// TIA Portal project "btl" (V17)

(* hardware
DEVICE "S7-1200 station_1"  S7-1200 Station
   slot 0: "Rack_0"  S7-1200 Rack  Rack  V1.0
   slot 1: "PLC_1"  CPU 1215C DC/DC/DC  6ES7 215-1AG40-0XB0  V4.5
   slot 2: "DI 16/DQ 16x24VDC SINK_1"  SM 1223 DI16/DQ16 x 24VDC SINK  6ES7 223-1BL32-1XB0  V2.0
   slot 3: "AI 8x13BIT_1"  6ES7 231-4HF32-0XB0  V2.1
   slot 4: "DI 8x24VDC_1"  SM 1221 DI8 x 24VDC  6ES7 221-1BF30-0XB0  V1.0
DEVICE "PC-System_1"  SIMATIC PC station
   slot 0: "SIMATIC PC station"  Rail  SIMATIC PC-Station  V1.0
      slot 125: "Stationmanager"  Station_Manager  V6.0.4
   slot 1: "HMI_RT_1"  WinCC RT Advanced  6AV2 104-0xxxx-xxxx  17.0.0.0
      slot 33792: "Computer interface"  Host interface
   slot 2: "IE general_1"  IE General  IE_CP  V8.2.0
      slot 1: "PROFINET interface"  IEGeneral.Interface.8.2.0
*)

// ===== PLC "PLC_1"  CPU 1215C DC/DC/DC =====

VAR_GLOBAL   // PLC tag table "Default tag table"
   "System_Byte" AT %MB1 : Byte;
   "FirstScan" AT %M1.0 : Bool;
   "DiagStatusUpdate" AT %M1.1 : Bool;
   "AlwaysTRUE" AT %M1.2 : Bool;
   "AlwaysFALSE" AT %M1.3 : Bool;
   "Clock_Byte" AT %MB0 : Byte;
   "Clock_10Hz" AT %M0.0 : Bool;
   "Clock_5Hz" AT %M0.1 : Bool;
   "Clock_2.5Hz" AT %M0.2 : Bool;
   "Clock_2Hz" AT %M0.3 : Bool;
   "Clock_1.25Hz" AT %M0.4 : Bool;
   "Clock_1Hz" AT %M0.5 : Bool;
   "Clock_0.625Hz" AT %M0.6 : Bool;
   "Clock_0.5Hz" AT %M0.7 : Bool;
END_VAR

VAR_GLOBAL   // PLC tag table "CB_analog"
   "I_Can_huong" AT %IW64 : Int;
   "I_can_mau" AT %IW66 : Int;
   "I_can_Duong" AT %IW68 : Int;
   "I_can_nuoc_TRON" AT %IW70 : Int;
   "I_Can_nuoc_xuc_khi" AT %IW72 : Int;
   "I_Can_PG" AT %IW74 : Int;
   "I_Can_CO2" AT %IW76 : Int;
   "I_bon_1" AT %IW82 : Int;
   "I_bon_2" AT %IW84 : Int;
   "I_bon_3" AT %IW86 : Int;
END_VAR

VAR_GLOBAL   // PLC tag table "INPUT_I"
   "I_mode" AT %I0.0 : Bool;
   "I_start" AT %I0.1 : Bool;
   "I_Stop" AT %I0.2 : Bool;
   "I_SW_V1_Huong" AT %I0.3 : Bool;
   "I_SW_V2_Huong" AT %I0.4 : Bool;
   "I_SW_V1_mau" AT %I0.5 : Bool;
   "I_SW_V2_mau" AT %I0.6 : Bool;
   "I_SW_V1_PG" AT %I0.7 : Bool;
   "I_SW_V2_PG" AT %I1.0 : Bool;
   "I_SW_V1_Duong" AT %I1.1 : Bool;
   "I_SW_V2_Duong" AT %I1.2 : Bool;
   "I_SW_V1_Nuoc_Tron" AT %I1.3 : Bool;
   "I_SW_V2_Nuoc_Tron" AT %I1.4 : Bool;
   "I_SW_V1_Nuoc_Xuc_Khi" AT %I1.5 : Bool;
   "I_SW_V2_Nuoc_Xuc_Khi" AT %I1.6 : Bool;
   "I_SW_V1_CO2" AT %I1.7 : Bool;
   "I_SW_V2_CO2" AT %I2.0 : Bool;
   "I_SW_BOM_TRON" AT %I2.1 : Bool;
   "I_SW_LAM_LANH" AT %I2.2 : Bool;
   "I_SW_BOM_1" AT %I2.3 : Bool;
   "I_SW_BOM_2" AT %I2.4 : Bool;
   "I_SW_LO_DOT" AT %I2.5 : Bool;
   "I_SW_VAN_XA" AT %I2.6 : Bool;
   "I_SW_BANG_TAI" AT %I2.7 : Bool;
   "I_CB_LOW_HUONG" AT %I3.0 : Bool;
   "I_CB_LOW_MAU" AT %I3.1 : Bool;
   "I_CB_LOW_PG" AT %I3.2 : Bool;
   "I_CB_LOW_DUONG" AT %I3.3 : Bool;
   "I_CB_LOW_NUOC" AT %I3.4 : Bool;
   "I_CB_LOW_CO2" AT %I3.5 : Bool;
   "I_CB_CHAI" AT %I3.6 : Bool;
END_VAR

VAR_GLOBAL   // PLC tag table "INPUT_M"
   "M_mode" AT %M10.0 : Bool;
   "M_start" AT %M10.1 : Bool;
   "M_Stop" AT %M10.2 : Bool;
   "M_SW_V1_Huong" AT %M10.3 : Bool;
   "M_SW_V2_Huong" AT %M10.4 : Bool;
   "M_SW_V1_mau" AT %M10.5 : Bool;
   "M_SW_V2_mau" AT %M10.6 : Bool;
   "M_SW_V1_PG" AT %M10.7 : Bool;
   "M_SW_V2_PG" AT %M11.0 : Bool;
   "M_SW_V1_Duong" AT %M11.1 : Bool;
   "M_SW_V2_Duong" AT %M11.2 : Bool;
   "M_SW_V1_Nuoc_Tron" AT %M11.3 : Bool;
   "M_SW_V2_Nuoc_Tron" AT %M11.4 : Bool;
   "M_SW_V1_Nuoc_Xuc_Khi" AT %M11.5 : Bool;
   "M_SW_V2_Nuoc_Xuc_Khi" AT %M11.6 : Bool;
   "M_SW_V1_CO2" AT %M11.7 : Bool;
   "M_SW_V2_CO2" AT %M12.0 : Bool;
   "M_SW_BOM_TRON" AT %M12.1 : Bool;
   "M_SW_LAM_LANH" AT %M12.2 : Bool;
   "M_SW_BOM_1" AT %M12.3 : Bool;
   "M_SW_BOM_2" AT %M12.4 : Bool;
   "M_SW_LO_DOT" AT %M12.5 : Bool;
   "M_SW_VAN_XA" AT %M12.6 : Bool;
   "M_SW_BANG_TAI" AT %M12.7 : Bool;
   "M_CB_LOW_HUONG" AT %M13.0 : Bool;
   "M_CB_LOW_MAU" AT %M13.1 : Bool;
   "M_CB_LOW_PG" AT %M13.2 : Bool;
   "M_CB_LOW_DUONG" AT %M13.3 : Bool;
   "M_CB_LOW_NUOC" AT %M13.4 : Bool;
   "M_CB_LOW_CO2" AT %MD500 : Real;
   "M_CB_LOW_BON_2" AT %MD504 : Real;
   "M_CB_CHAI" AT %M13.7 : Bool;
END_VAR

VAR_GLOBAL   // PLC tag table "OUTPUT"
   "Q_den_Auto" AT %Q0.0 : Bool;
   "Q_Den_Manual" AT %Q0.1 : Bool;
   "Q_Den_loi" AT %Q0.2 : Bool;
   "Q_V1_Huong" AT %Q0.3 : Bool;
   "Q_V2_Huong" AT %Q0.4 : Bool;
   "Q_V1_Mau" AT %Q0.5 : Bool;
   "Q_V2_Mau" AT %Q0.6 : Bool;
   "Q_V1_PG" AT %Q0.7 : Bool;
   "Q_V2_PG" AT %Q1.0 : Bool;
   "Q_V1_Nuoc_Tron" AT %Q1.1 : Bool;
   "Q_V2_Nuoc_tron" AT %Q1.2 : Bool;
   "Q_V1_Duong" AT %Q1.3 : Bool;
   "Q_V2_Duong" AT %Q1.4 : Bool;
   "Q_V1_Nuoc_Khi" AT %Q1.5 : Bool;
   "Q_V2_Xuc_Khi" AT %Q1.6 : Bool;
   "Q_V1_CO2" AT %Q1.7 : Bool;
   "Q_V2_CO2" AT %Q2.0 : Bool;
   "Q_BOM_TRON" AT %Q2.1 : Bool;
   "Q_LAM_LANH" AT %Q2.2 : Bool;
   "Q_BOM_1" AT %Q2.3 : Bool;
   "Q_BOM_2" AT %Q2.4 : Bool;
   "Q_VAN_XA" AT %Q2.5 : Bool;
   "Q_LO_DOT" AT %Q2.6 : Bool;
   "Q_BT" AT %Q2.7 : Bool;
END_VAR

VAR_GLOBAL   // PLC tag table "OUTPUT_AUTO"
   "Q_AUTO_den_Auto" AT %M20.0 : Bool;
   "Q_AUTO_Den_Manual" AT %M20.1 : Bool;
   "Q_AUTO_Den_loi" AT %M20.2 : Bool;
   "Q_AUTO_V1_Huong" AT %M20.3 : Bool;
   "Q_AUTO_V2_Huong" AT %M20.4 : Bool;
   "Q_AUTO_V1_Mau" AT %M20.5 : Bool;
   "Q_AUTO_V2_Mau" AT %M20.6 : Bool;
   "Q_AUTO_V1_PG" AT %M20.7 : Bool;
   "Q_AUTO_V2_PG" AT %M21.0 : Bool;
   "Q_AUTO_V1_Nuoc_Tron" AT %M21.1 : Bool;
   "Q_AUTO_V2_Nuoc_tron" AT %M21.2 : Bool;
   "Q_AUTO_V1_Duong" AT %M21.3 : Bool;
   "Q_AUTO_V2_Duong" AT %M21.4 : Bool;
   "Q_AUTO_V1_Nuoc_Khi" AT %M21.5 : Bool;
   "Q_AUTO_V2_Xuc_Khi" AT %M21.6 : Bool;
   "Q_AUTO_V1_CO2" AT %M21.7 : Bool;
   "Q_AUTO_V2_CO2" AT %M22.0 : Bool;
   "Q_AUTO_BOM_TRON" AT %M22.1 : Bool;
   "Q_AUTO_LAM_LANH" AT %M22.2 : Bool;
   "Q_AUTO_BOM_1" AT %M22.3 : Bool;
   "Q_AUTO_BOM_2" AT %M22.4 : Bool;
   "Q_AUTO_VAN_XA" AT %M22.5 : Bool;
   "Q_AUTO_LO_DOT" AT %M22.6 : Bool;
   "Q_AUTO_BT" AT %M22.7 : Bool;
END_VAR

VAR_GLOBAL   // PLC tag table "OUTPUT_MANUAL"
   "Q_MAN_den_Auto" AT %M30.0 : Bool;
   "Q_MAN_Den_Manual" AT %M30.1 : Bool;
   "Q_MAN_Den_loi" AT %M30.2 : Bool;
   "Q_MAN_V1_Huong" AT %M30.3 : Bool;
   "Q_MAN_V2_Huong" AT %M30.4 : Bool;
   "Q_MAN_V1_Mau" AT %M30.5 : Bool;
   "Q_MAN_V2_Mau" AT %M30.6 : Bool;
   "Q_MAN_V1_PG" AT %M30.7 : Bool;
   "Q_MAN_V2_PG" AT %M31.0 : Bool;
   "Q_MAN_V1_Nuoc_Tron" AT %M31.1 : Bool;
   "Q_MAN_V2_Nuoc_tron" AT %M31.2 : Bool;
   "Q_MAN_V1_Duong" AT %M31.3 : Bool;
   "Q_MAN_V2_Duong" AT %M31.4 : Bool;
   "Q_MAN_V1_Nuoc_Khi" AT %M31.5 : Bool;
   "Q_MAN_V2_Xuc_Khi" AT %M31.6 : Bool;
   "Q_MAN_V1_CO2" AT %M31.7 : Bool;
   "Q_MAN_V2_CO2" AT %M32.0 : Bool;
   "Q_MAN_BOM_TRON" AT %M32.1 : Bool;
   "Q_MAN_LAM_LANH" AT %M32.2 : Bool;
   "Q_MAN_BOM_1" AT %M32.3 : Bool;
   "Q_MAN_BOM_2" AT %M32.4 : Bool;
   "Q_MAN_VAN_XA" AT %M32.5 : Bool;
   "Q_MAN_LO_DOT" AT %M32.6 : Bool;
   "Q_MAN_BT" AT %M32.7 : Bool;
END_VAR

VAR_GLOBAL   // PLC tag table "GT_Thuc_TE"
   "Act_time_Khuay" AT %MW400 : Int;
   "Act_nhiet_do" AT %MD402 : Real;
   "Act_me" AT %MW406 : Int;
   "Act_can_huong" AT %MD408 : Real;
   "Act_can_mau" AT %MD412 : Real;
   "Act_can_duong" AT %MD416 : Real;
   "Act_can_PG" AT %MD420 : Real;
   "Act_can_nuoc_tron" AT %MD424 : Real;
   "Act_can_nuoc_xuc_khi" AT %MD428 : Real;
   "Act_Can_CO2" AT %MD432 : Real;
   "Act_So_chai" AT %MW436 : Int;
   "Act_bon_1" AT %MD440 : Real;
   "Act_bon_2" AT %MD444 : Real;
   "Act_bon_3" AT %MD448 : Real;
END_VAR

VAR_GLOBAL   // PLC tag table "Trung_gian"
   "TG_Button_Simulation" AT %M40.0 : Bool;
   "TG_Step_1" AT %M40.1 : Bool;
   "TG_Step_2" AT %M40.2 : Bool;
   "TG_Step_3" AT %M40.3 : Bool;
   "TG_Step_4" AT %M40.4 : Bool;
   "TG_Step_5" AT %M40.5 : Bool;
   "TG_Step_6" AT %M40.6 : Bool;
   "TG_Step_7" AT %M40.7 : Bool;
   "TG_DK_RUN" AT %M41.0 : Bool;
   "TG_Lap_lai" AT %M41.1 : Bool;
   "TG_Can_Xong_huong" AT %M41.2 : Bool;
   "TG_Xung_100ms" AT %M41.3 : Bool;
   "TG_Can_Xong_mau" AT %M41.4 : Bool;
   "TG_Can_Xong_PG" AT %M41.5 : Bool;
   "TG_can_Xong_Nuoc_Khi" AT %M41.6 : Bool;
   "TG_Can_Xong_CO2" AT %M41.7 : Bool;
   "TG_xong_nuoc_tron" AT %M42.0 : Bool;
   "TG_Xong_Nuoc_khi" AT %M42.1 : Bool;
   "TG_xong_huong" AT %M42.2 : Bool;
   "TG_Xong_mau" AT %M42.3 : Bool;
   "TG_Xong_PG" AT %M42.4 : Bool;
   "TG_Xong_duong" AT %M42.5 : Bool;
   "TG_Xong_CO2" AT %M42.6 : Bool;
   "TG_Xong_Khuay" AT %M42.7 : Bool;
   "TG_Xong_Dot" AT %M43.0 : Bool;
   "TG_Thoi_Gian_Dong_SP" AT %M43.1 : Bool;
   "TG_XONG_BANG_TAI" AT %M43.2 : Bool;
   "TG_DONE_CHU_TRINH" AT %M43.3 : Bool;
   "TG_VT_SP" AT %MD508 : DInt;
   "TG_TG_SP" AT %MD512 : DInt;
   "TG_Can_huong" AT %MD516 : Real;
   "TG_Can_mau" AT %MD520 : Real;
   "TG_Can_PG" AT %MD524 : Real;
   "TG_CAn_Duong" AT %MD528 : Real;
   "TG_Can_nuoc_tron" AT %MD532 : Real;
   "TG_Can_nuoc_khi" AT %MD536 : Real;
   "TG_Can_CO2" AT %MD540 : Real;
   "TG_BON1" AT %M43.4 : Bool;
   "TG_BON2" AT %M43.5 : Bool;
   "TG_BON3" AT %M43.6 : Bool;
   "TG_V_BON1" AT %MD544 : Real;
   "TG_V_BON2" AT %MD548 : Real;
   "TG_V_BON3" AT %MD552 : Real;
   "TG_LO_DOT" AT %M43.7 : Bool;
END_VAR

VAR_GLOBAL   // PLC tag table "Trung_giang_Xung"
   "P1" AT %M50.0 : Bool;
   "P2" AT %M50.1 : Bool;
   "P3" AT %M50.2 : Bool;
   "P4" AT %M50.3 : Bool;
   "P5" AT %M50.4 : Bool;
   "P6" AT %M50.5 : Bool;
   "P7" AT %M50.6 : Bool;
   "P8" AT %M50.7 : Bool;
   "P9" AT %M51.0 : Bool;
   "P10" AT %M51.1 : Bool;
   "P11" AT %M51.2 : Bool;
   "P12" AT %M51.3 : Bool;
   "P13" AT %M51.4 : Bool;
   "P14" AT %M51.5 : Bool;
   "P15" AT %M51.6 : Bool;
   "P16" AT %M51.7 : Bool;
   "P17" AT %M52.0 : Bool;
   "P18" AT %M52.1 : Bool;
   "P19" AT %M52.2 : Bool;
   "P20" AT %M52.3 : Bool;
   "P21" AT %M52.4 : Bool;
   "P22" AT %M52.5 : Bool;
   "P23" AT %M52.6 : Bool;
   "P24" AT %M52.7 : Bool;
   "P25" AT %M53.0 : Bool;
   "P26" AT %M53.1 : Bool;
   "P27" AT %M53.2 : Bool;
   "P28" AT %M53.3 : Bool;
   "P29" AT %M53.4 : Bool;
   "P30" AT %M53.5 : Bool;
   "P31" AT %M53.6 : Bool;
   "P32" AT %M53.7 : Bool;
   "P33" AT %M54.0 : Bool;
   "P34" AT %M54.1 : Bool;
   "P35" AT %M54.2 : Bool;
   "P36" AT %M54.3 : Bool;
   "P37" AT %M54.4 : Bool;
   "P38" AT %M54.5 : Bool;
   "P39" AT %M54.6 : Bool;
   "P40" AT %M54.7 : Bool;
   "P41" AT %M55.0 : Bool;
   "P42" AT %M55.1 : Bool;
END_VAR

VAR_GLOBAL   // PLC tag table "Setting"
   "Set_can_huong" AT %MD200 : Real;
   "Set_can_mau" AT %MD204 : Real;
   "Set_can_PG" AT %MD208 : Real;
   "Set_can_Duong" AT %MD212 : Real;
   "Set_Can_nuoc_Tron" AT %MD216 : Real;
   "Set_Can_nuoc_xuc_khi" AT %MD220 : Real;
   "Set_Can_CO2" AT %MD224 : Real;
   "Set_thoi_gian_khuay" AT %MW228 : Int;
   "Set_nhiet_do" AT %MD300 : Real;
   "Set_me_tron" AT %MW304 : Int;
END_VAR

VAR_GLOBAL   // PLC tag table "TRONG LUONG DAT DUOC"
   "TL_Huong" AT %MD600 : Real;
   "TL_mau" AT %MD604 : Real;
   "TL_Duong" AT %MD608 : Real;
   "TL_PG" AT %MD612 : Real;
   "TL_nuoc_tron" AT %MD616 : Real;
   "TL_CO2" AT %MD620 : Real;
   "TL_Nuoc_KHi" AT %MD624 : Real;
   "TL_San_Pham" AT %MD628 : Real;
   "TL_thoiGian_khuay" AT %MD632 : DInt;
   "TL_nhietdo" AT %MD636 : Real;
END_VAR

// folder: System blocks/Program resources

DATA_BLOCK "IEC_Timer_0_DB"   // DB1
{ S7_Optimized_Access := 'TRUE' }
AUTHOR : Simatic
FAMILY : IEC
NAME : IEC_TMR
VERSION : 1.0
// stored: InstanceOfName IEC_TIMER
"IEC_TIMER"
BEGIN
END_DATA_BLOCK

DATA_BLOCK "IEC_Timer_0_DB_1"   // DB2
{ S7_Optimized_Access := 'TRUE' }
AUTHOR : Simatic
FAMILY : IEC
NAME : IEC_TMR
VERSION : 1.0
// stored: InstanceOfName IEC_TIMER
"IEC_TIMER"
BEGIN
END_DATA_BLOCK

DATA_BLOCK "IEC_Timer_0_DB_2"   // DB3
{ S7_Optimized_Access := 'TRUE' }
AUTHOR : Simatic
FAMILY : IEC
NAME : IEC_TMR
VERSION : 1.0
// stored: InstanceOfName IEC_TIMER
"IEC_TIMER"
BEGIN
END_DATA_BLOCK

DATA_BLOCK "IEC_Timer_0_DB_3"   // DB4
{ S7_Optimized_Access := 'TRUE' }
AUTHOR : Simatic
FAMILY : IEC
NAME : IEC_TMR
VERSION : 1.0
// stored: InstanceOfName IEC_TIMER
"IEC_TIMER"
BEGIN
END_DATA_BLOCK

// folder: (top level)

FUNCTION "FC_ANALOG" : Void   // FC1, LAD
{ S7_Optimized_Access := 'TRUE' }
VERSION : 0.1
BEGIN

REGION Network 1: Can Huong
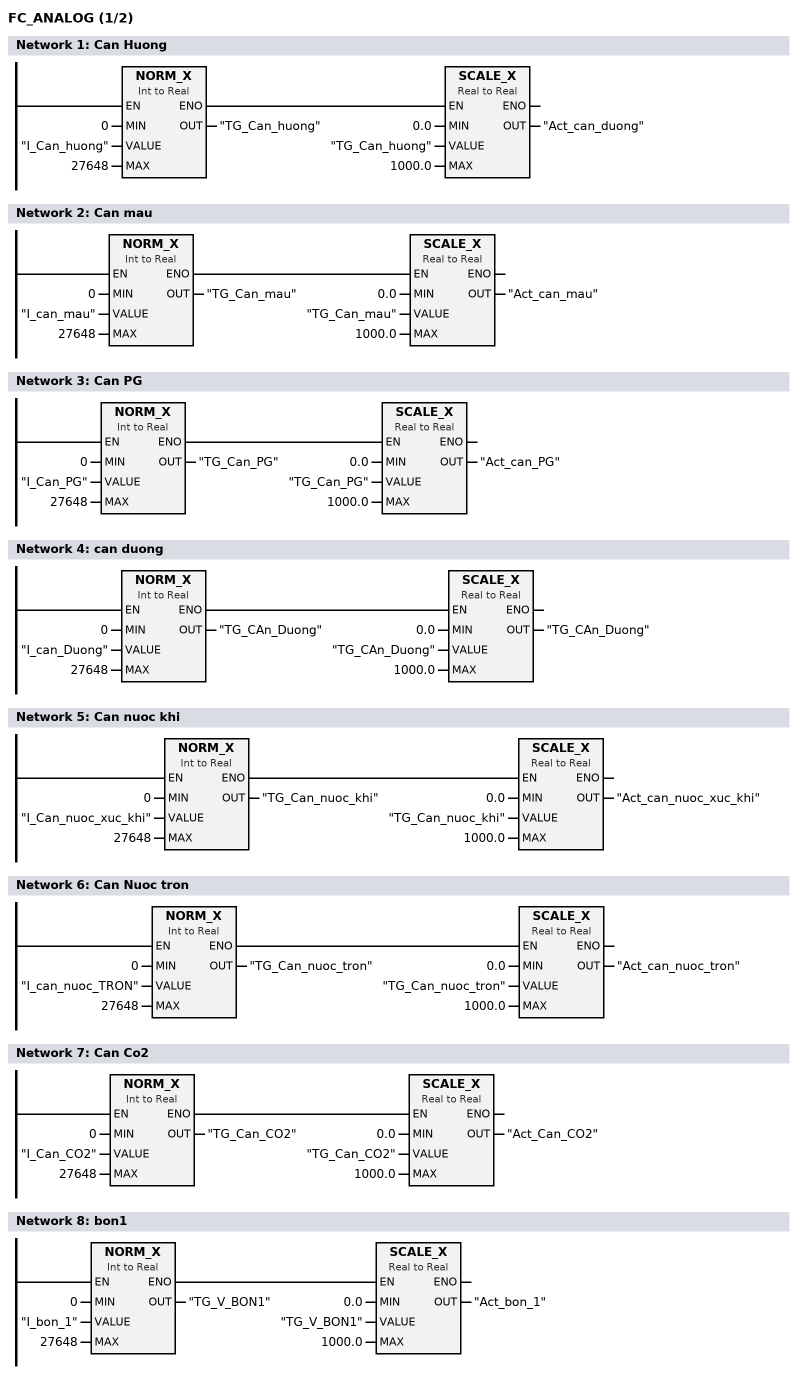
   RUNG wire#powerrail
      { S7_Templates := "[SrcType := Int, DestType := Real]" } Normalize(min := 0, value := "I_Can_huong", max := 27648, out => "TG_Can_huong")
      { S7_Templates := "[SrcType := Real, DestType := Real]" } Scale(min := 0.0, value := "TG_Can_huong", max := 1000.0, out => "Act_can_duong")
   END_RUNG
   // the same network as SCL:
   "TG_Can_huong" := NORM_X(MIN := 0, VALUE := "I_Can_huong", MAX := 27648);
   "Act_can_duong" := SCALE_X(MIN := 0.0, VALUE := "TG_Can_huong", MAX := 1000.0);
END_REGION

REGION Network 2: Can mau
   RUNG wire#powerrail
      { S7_Templates := "[SrcType := Int, DestType := Real]" } Normalize(min := 0, value := "I_can_mau", max := 27648, out => "TG_Can_mau")
      { S7_Templates := "[SrcType := Real, DestType := Real]" } Scale(min := 0.0, value := "TG_Can_mau", max := 1000.0, out => "Act_can_mau")
   END_RUNG
   // the same network as SCL:
   "TG_Can_mau" := NORM_X(MIN := 0, VALUE := "I_can_mau", MAX := 27648);
   "Act_can_mau" := SCALE_X(MIN := 0.0, VALUE := "TG_Can_mau", MAX := 1000.0);
END_REGION

REGION Network 3: Can PG
   RUNG wire#powerrail
      { S7_Templates := "[SrcType := Int, DestType := Real]" } Normalize(min := 0, value := "I_Can_PG", max := 27648, out => "TG_Can_PG")
      { S7_Templates := "[SrcType := Real, DestType := Real]" } Scale(min := 0.0, value := "TG_Can_PG", max := 1000.0, out => "Act_can_PG")
   END_RUNG
   // the same network as SCL:
   "TG_Can_PG" := NORM_X(MIN := 0, VALUE := "I_Can_PG", MAX := 27648);
   "Act_can_PG" := SCALE_X(MIN := 0.0, VALUE := "TG_Can_PG", MAX := 1000.0);
END_REGION

REGION Network 4: can duong
   RUNG wire#powerrail
      { S7_Templates := "[SrcType := Int, DestType := Real]" } Normalize(min := 0, value := "I_can_Duong", max := 27648, out => "TG_CAn_Duong")
      { S7_Templates := "[SrcType := Real, DestType := Real]" } Scale(min := 0.0, value := "TG_CAn_Duong", max := 1000.0, out => "TG_CAn_Duong")
   END_RUNG
   // the same network as SCL:
   "TG_CAn_Duong" := NORM_X(MIN := 0, VALUE := "I_can_Duong", MAX := 27648);
   "TG_CAn_Duong" := SCALE_X(MIN := 0.0, VALUE := "TG_CAn_Duong", MAX := 1000.0);
END_REGION

REGION Network 5: Can nuoc khi
   RUNG wire#powerrail
      { S7_Templates := "[SrcType := Int, DestType := Real]" } Normalize(min := 0, value := "I_Can_nuoc_xuc_khi", max := 27648, out => "TG_Can_nuoc_khi")
      { S7_Templates := "[SrcType := Real, DestType := Real]" } Scale(min := 0.0, value := "TG_Can_nuoc_khi", max := 1000.0, out => "Act_can_nuoc_xuc_khi")
   END_RUNG
   // the same network as SCL:
   "TG_Can_nuoc_khi" := NORM_X(MIN := 0, VALUE := "I_Can_nuoc_xuc_khi", MAX := 27648);
   "Act_can_nuoc_xuc_khi" := SCALE_X(MIN := 0.0, VALUE := "TG_Can_nuoc_khi", MAX := 1000.0);
END_REGION

REGION Network 6: Can Nuoc tron
   RUNG wire#powerrail
      { S7_Templates := "[SrcType := Int, DestType := Real]" } Normalize(min := 0, value := "I_can_nuoc_TRON", max := 27648, out => "TG_Can_nuoc_tron")
      { S7_Templates := "[SrcType := Real, DestType := Real]" } Scale(min := 0.0, value := "TG_Can_nuoc_tron", max := 1000.0, out => "Act_can_nuoc_tron")
   END_RUNG
   // the same network as SCL:
   "TG_Can_nuoc_tron" := NORM_X(MIN := 0, VALUE := "I_can_nuoc_TRON", MAX := 27648);
   "Act_can_nuoc_tron" := SCALE_X(MIN := 0.0, VALUE := "TG_Can_nuoc_tron", MAX := 1000.0);
END_REGION

REGION Network 7: Can Co2
   RUNG wire#powerrail
      { S7_Templates := "[SrcType := Int, DestType := Real]" } Normalize(min := 0, value := "I_Can_CO2", max := 27648, out => "TG_Can_CO2")
      { S7_Templates := "[SrcType := Real, DestType := Real]" } Scale(min := 0.0, value := "TG_Can_CO2", max := 1000.0, out => "Act_Can_CO2")
   END_RUNG
   // the same network as SCL:
   "TG_Can_CO2" := NORM_X(MIN := 0, VALUE := "I_Can_CO2", MAX := 27648);
   "Act_Can_CO2" := SCALE_X(MIN := 0.0, VALUE := "TG_Can_CO2", MAX := 1000.0);
END_REGION

REGION Network 8: bon1
   RUNG wire#powerrail
      { S7_Templates := "[SrcType := Int, DestType := Real]" } Normalize(min := 0, value := "I_bon_1", max := 27648, out => "TG_V_BON1")
      { S7_Templates := "[SrcType := Real, DestType := Real]" } Scale(min := 0.0, value := "TG_V_BON1", max := 1000.0, out => "Act_bon_1")
   END_RUNG
   // the same network as SCL:
   "TG_V_BON1" := NORM_X(MIN := 0, VALUE := "I_bon_1", MAX := 27648);
   "Act_bon_1" := SCALE_X(MIN := 0.0, VALUE := "TG_V_BON1", MAX := 1000.0);
END_REGION

REGION Network 9: bon2
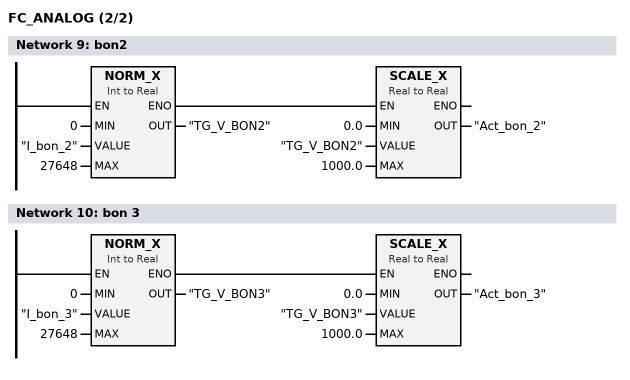
   RUNG wire#powerrail
      { S7_Templates := "[SrcType := Int, DestType := Real]" } Normalize(min := 0, value := "I_bon_2", max := 27648, out => "TG_V_BON2")
      { S7_Templates := "[SrcType := Real, DestType := Real]" } Scale(min := 0.0, value := "TG_V_BON2", max := 1000.0, out => "Act_bon_2")
   END_RUNG
   // the same network as SCL:
   "TG_V_BON2" := NORM_X(MIN := 0, VALUE := "I_bon_2", MAX := 27648);
   "Act_bon_2" := SCALE_X(MIN := 0.0, VALUE := "TG_V_BON2", MAX := 1000.0);
END_REGION

REGION Network 10: bon 3
   RUNG wire#powerrail
      { S7_Templates := "[SrcType := Int, DestType := Real]" } Normalize(min := 0, value := "I_bon_3", max := 27648, out => "TG_V_BON3")
      { S7_Templates := "[SrcType := Real, DestType := Real]" } Scale(min := 0.0, value := "TG_V_BON3", max := 1000.0, out => "Act_bon_3")
   END_RUNG
   // the same network as SCL:
   "TG_V_BON3" := NORM_X(MIN := 0, VALUE := "I_bon_3", MAX := 27648);
   "Act_bon_3" := SCALE_X(MIN := 0.0, VALUE := "TG_V_BON3", MAX := 1000.0);
END_REGION
END_FUNCTION

FUNCTION "FC_AUTO" : Void   // FC2, LAD
{ S7_Optimized_Access := 'TRUE' }
VERSION : 0.1
   VAR_TEMP   // added for the SCL form of the ladder/FBD networks
      _w1 : Bool;
      _w2 : Bool;
      _w3 : Bool;
      _w4 : Bool;
      _w5 : Bool;
      _w6 : Bool;
      _w7 : Bool;
      _w8 : Bool;
      _w9 : Bool;
      _w10 : Bool;
      _w11 : Bool;
      _w12 : Bool;
      _w13 : Bool;
      _w14 : Bool;
      _w15 : Bool;
      _w16 : Bool;
      _w17 : Bool;
      _w18 : Bool;
      _w19 : Bool;
      _w20 : Bool;
      _w21 : Bool;
   END_VAR
BEGIN

REGION Network 1: Điều Kiện Vận Hành
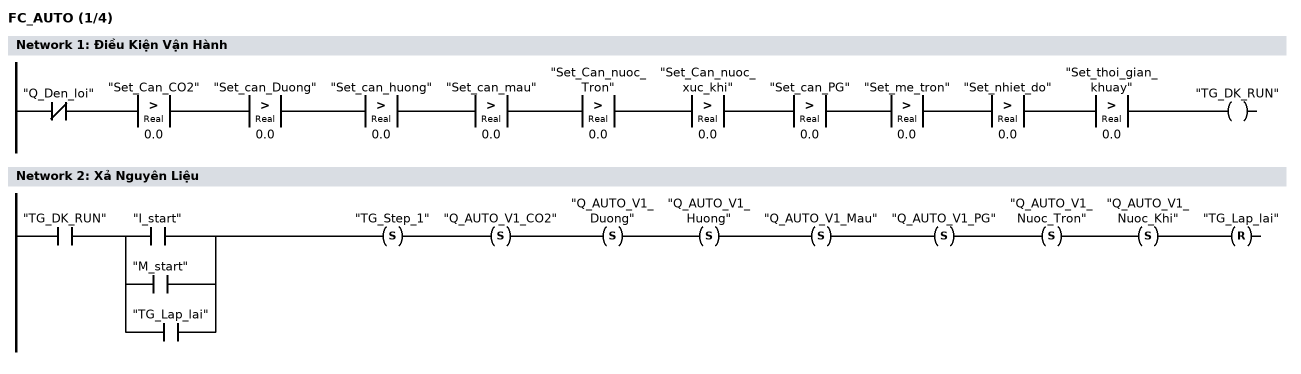
   RUNG wire#powerrail
      I_Contact( "Q_Den_loi" )
      { S7_Templates := "SrcType := Real" } GT_Contact(in1 := "Set_Can_CO2", in2 := 0.0)
      { S7_Templates := "SrcType := Real" } GT_Contact(in1 := "Set_can_Duong", in2 := 0.0)
      { S7_Templates := "SrcType := Real" } GT_Contact(in1 := "Set_can_huong", in2 := 0.0)
      { S7_Templates := "SrcType := Real" } GT_Contact(in1 := "Set_can_mau", in2 := 0.0)
      { S7_Templates := "SrcType := Real" } GT_Contact(in1 := "Set_Can_nuoc_Tron", in2 := 0.0)
      { S7_Templates := "SrcType := Real" } GT_Contact(in1 := "Set_Can_nuoc_xuc_khi", in2 := 0.0)
      { S7_Templates := "SrcType := Real" } GT_Contact(in1 := "Set_can_PG", in2 := 0.0)
      { S7_Templates := "SrcType := Real" } GT_Contact(in1 := "Set_me_tron", in2 := 0.0)
      { S7_Templates := "SrcType := Real" } GT_Contact(in1 := "Set_nhiet_do", in2 := 0.0)
      { S7_Templates := "SrcType := Real" } GT_Contact(in1 := "Set_thoi_gian_khuay", in2 := 0.0)
      Coil( "TG_DK_RUN" )
   END_RUNG
   // the same network as SCL:
   "TG_DK_RUN" := NOT "Q_Den_loi" AND ("Set_Can_CO2" > 0.0) AND ("Set_can_Duong" > 0.0) AND ("Set_can_huong" > 0.0) AND ("Set_can_mau" > 0.0) AND ("Set_Can_nuoc_Tron" > 0.0) AND ("Set_Can_nuoc_xuc_khi" > 0.0) AND ("Set_can_PG" > 0.0) AND ("Set_me_tron" > 0.0) AND ("Set_nhiet_do" > 0.0) AND ("Set_thoi_gian_khuay" > 0.0);
END_REGION

REGION Network 2: Xả Nguyên Liệu
   RUNG wire#powerrail
      Contact( "TG_DK_RUN" )
      wire#w1
      Contact( "I_start" )
      wire#w2
      S_Coil( "TG_Step_1" )
      S_Coil( "Q_AUTO_V1_CO2" )
      S_Coil( "Q_AUTO_V1_Duong" )
      S_Coil( "Q_AUTO_V1_Huong" )
      S_Coil( "Q_AUTO_V1_Mau" )
      S_Coil( "Q_AUTO_V1_PG" )
      S_Coil( "Q_AUTO_V1_Nuoc_Tron" )
      S_Coil( "Q_AUTO_V1_Nuoc_Khi" )
      R_Coil( "TG_Lap_lai" )
   END_RUNG
   RUNG wire#w1
      Contact( "M_start" )
   END_RUNG wire#w2
   RUNG wire#w1
      Contact( "TG_Lap_lai" )
   END_RUNG wire#w2
   // the same network as SCL:
   IF "TG_DK_RUN" AND ("I_start" OR "M_start" OR "TG_Lap_lai") THEN
       "TG_Step_1" := TRUE;
       "Q_AUTO_V1_CO2" := TRUE;
       "Q_AUTO_V1_Duong" := TRUE;
       "Q_AUTO_V1_Huong" := TRUE;
       "Q_AUTO_V1_Mau" := TRUE;
       "Q_AUTO_V1_PG" := TRUE;
       "Q_AUTO_V1_Nuoc_Tron" := TRUE;
       "Q_AUTO_V1_Nuoc_Khi" := TRUE;
       "TG_Lap_lai" := FALSE;
   END_IF;
END_REGION

REGION Network 3: Cân Hương, Đường, Màu , Phụ Gia , Nước , CO2
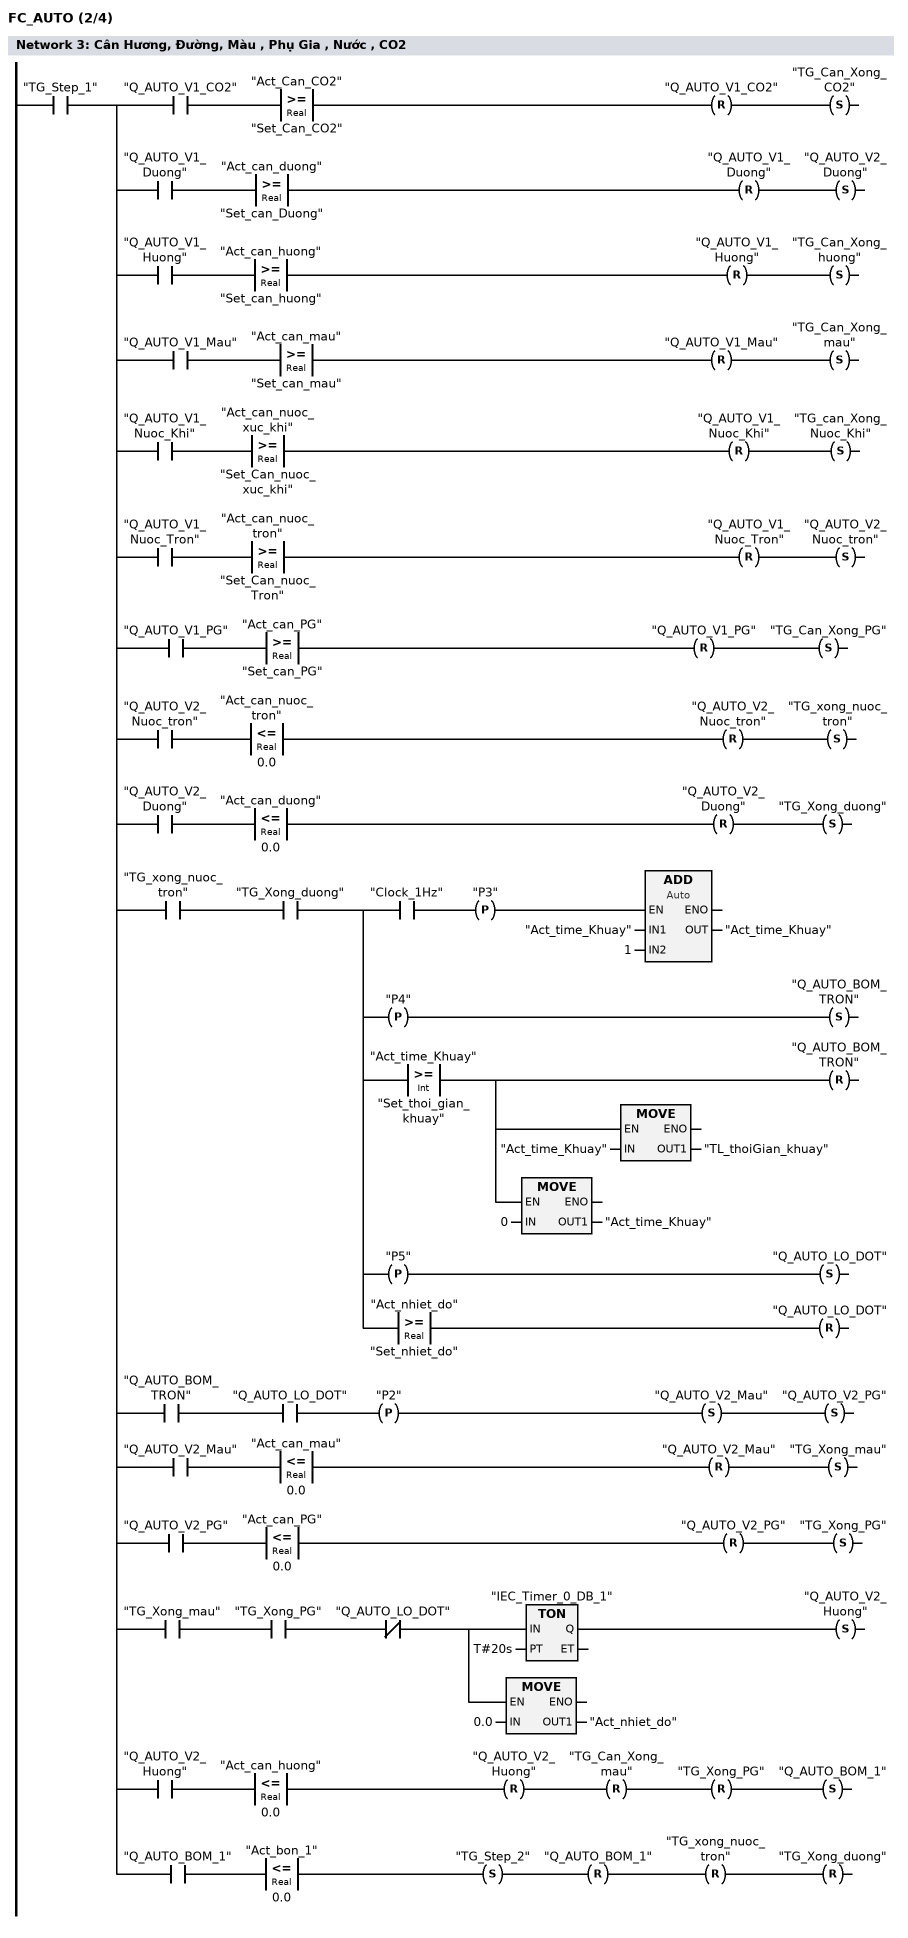
   #_w1 := "TG_Step_1" AND "Q_AUTO_V1_CO2" AND ("Act_Can_CO2" >= "Set_Can_CO2");
   IF #_w1 THEN
       "Q_AUTO_V1_CO2" := FALSE;
       "TG_Can_Xong_CO2" := TRUE;
   END_IF;
   #_w2 := "TG_Step_1" AND "Q_AUTO_V1_Duong" AND ("Act_can_duong" >= "Set_can_Duong");
   IF #_w2 THEN
       "Q_AUTO_V1_Duong" := FALSE;
       "Q_AUTO_V2_Duong" := TRUE;
   END_IF;
   #_w3 := "TG_Step_1" AND "Q_AUTO_V1_Huong" AND ("Act_can_huong" >= "Set_can_huong");
   IF #_w3 THEN
       "Q_AUTO_V1_Huong" := FALSE;
       "TG_Can_Xong_huong" := TRUE;
   END_IF;
   #_w4 := "TG_Step_1" AND "Q_AUTO_V1_Mau" AND ("Act_can_mau" >= "Set_can_mau");
   IF #_w4 THEN
       "Q_AUTO_V1_Mau" := FALSE;
       "TG_Can_Xong_mau" := TRUE;
   END_IF;
   #_w5 := "TG_Step_1" AND "Q_AUTO_V1_Nuoc_Khi" AND ("Act_can_nuoc_xuc_khi" >= "Set_Can_nuoc_xuc_khi");
   IF #_w5 THEN
       "Q_AUTO_V1_Nuoc_Khi" := FALSE;
       "TG_can_Xong_Nuoc_Khi" := TRUE;
   END_IF;
   #_w6 := "TG_Step_1" AND "Q_AUTO_V1_Nuoc_Tron" AND ("Act_can_nuoc_tron" >= "Set_Can_nuoc_Tron");
   IF #_w6 THEN
       "Q_AUTO_V1_Nuoc_Tron" := FALSE;
       "Q_AUTO_V2_Nuoc_tron" := TRUE;
   END_IF;
   #_w7 := "TG_Step_1" AND "Q_AUTO_V1_PG" AND ("Act_can_PG" >= "Set_can_PG");
   IF #_w7 THEN
       "Q_AUTO_V1_PG" := FALSE;
       "TG_Can_Xong_PG" := TRUE;
   END_IF;
   #_w8 := "TG_Step_1" AND "Q_AUTO_V2_Nuoc_tron" AND ("Act_can_nuoc_tron" <= 0.0);
   IF #_w8 THEN
       "Q_AUTO_V2_Nuoc_tron" := FALSE;
       "TG_xong_nuoc_tron" := TRUE;
   END_IF;
   #_w9 := "TG_Step_1" AND "Q_AUTO_V2_Duong" AND ("Act_can_duong" <= 0.0);
   IF #_w9 THEN
       "Q_AUTO_V2_Duong" := FALSE;
       "TG_Xong_duong" := TRUE;
   END_IF;
   #_w10 := "TG_Step_1" AND "TG_xong_nuoc_tron" AND "TG_Xong_duong";
   #_w11 := #_w10 AND "Clock_1Hz";
   #_w12 := #_w11 AND NOT "P3";   // rising edge
   "P3" := #_w11;
   IF #_w12 THEN "Act_time_Khuay" := "Act_time_Khuay" + 1; END_IF;
   #_w13 := #_w10 AND NOT "P4";   // rising edge
   "P4" := #_w10;
   IF #_w13 THEN "Q_AUTO_BOM_TRON" := TRUE; END_IF;
   IF #_w10 AND ("Act_time_Khuay" >= "Set_thoi_gian_khuay") THEN
       "Q_AUTO_BOM_TRON" := FALSE;
       "TL_thoiGian_khuay" := "Act_time_Khuay";
       "Act_time_Khuay" := 0;
   END_IF;
   #_w14 := #_w10 AND NOT "P5";   // rising edge
   "P5" := #_w10;
   IF #_w14 THEN "Q_AUTO_LO_DOT" := TRUE; END_IF;
   IF #_w10 AND ("Act_nhiet_do" >= "Set_nhiet_do") THEN "Q_AUTO_LO_DOT" := FALSE; END_IF;
   #_w15 := "TG_Step_1" AND "Q_AUTO_BOM_TRON" AND "Q_AUTO_LO_DOT";
   #_w16 := #_w15 AND NOT "P2";   // rising edge
   "P2" := #_w15;
   IF #_w16 THEN
       "Q_AUTO_V2_Mau" := TRUE;
       "Q_AUTO_V2_PG" := TRUE;
   END_IF;
   #_w17 := "TG_Step_1" AND "Q_AUTO_V2_Mau" AND ("Act_can_mau" <= 0.0);
   IF #_w17 THEN
       "Q_AUTO_V2_Mau" := FALSE;
       "TG_Xong_mau" := TRUE;
   END_IF;
   #_w18 := "TG_Step_1" AND "Q_AUTO_V2_PG" AND ("Act_can_PG" <= 0.0);
   IF #_w18 THEN
       "Q_AUTO_V2_PG" := FALSE;
       "TG_Xong_PG" := TRUE;
   END_IF;
   #_w19 := "TG_Step_1" AND "TG_Xong_mau" AND "TG_Xong_PG" AND NOT "Q_AUTO_LO_DOT";
   "IEC_Timer_0_DB_1".TON(IN := #_w19, PT := T#20s);
   IF "IEC_Timer_0_DB_1".Q THEN "Q_AUTO_V2_Huong" := TRUE; END_IF;
   IF #_w19 THEN "Act_nhiet_do" := 0.0; END_IF;
   #_w20 := "TG_Step_1" AND "Q_AUTO_V2_Huong" AND ("Act_can_huong" <= 0.0);
   IF #_w20 THEN
       "Q_AUTO_V2_Huong" := FALSE;
       "TG_Can_Xong_mau" := FALSE;
       "TG_Xong_PG" := FALSE;
       "Q_AUTO_BOM_1" := TRUE;
   END_IF;
   IF "TG_Step_1" AND "Q_AUTO_BOM_1" AND ("Act_bon_1" <= 0.0) THEN "TG_Step_2" := TRUE; END_IF;
   #_w21 := "TG_Step_1" AND "Q_AUTO_BOM_1" AND ("Act_bon_1" <= 0.0);
   IF #_w21 THEN
       "Q_AUTO_BOM_1" := FALSE;
       "TG_xong_nuoc_tron" := FALSE;
       "TG_Xong_duong" := FALSE;
   END_IF;
END_REGION

REGION Network 4
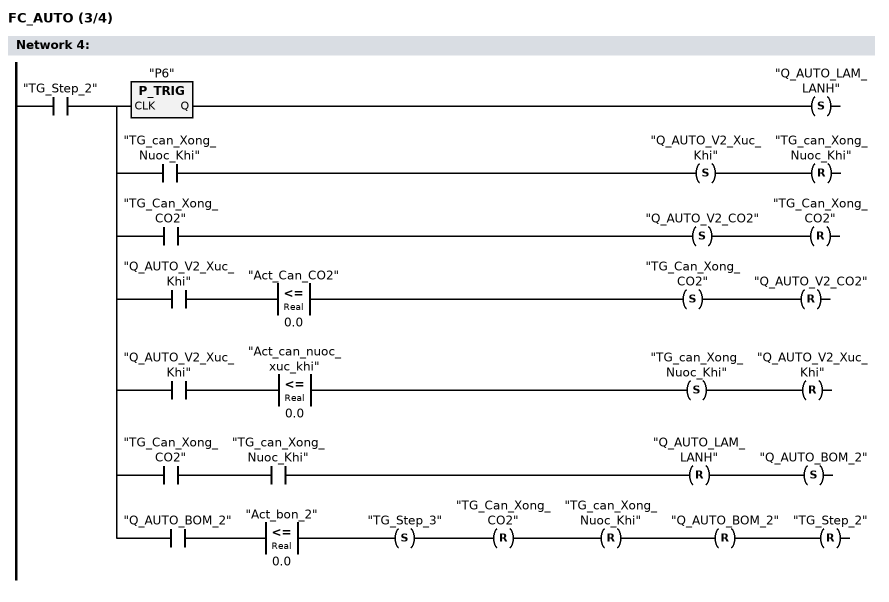
   RUNG wire#powerrail
      Contact( "TG_Step_2" )
      wire#w1
      P_Trig( "P6" )
      S_Coil( "Q_AUTO_LAM_LANH" )
   END_RUNG
   RUNG wire#w1
      Contact( "TG_can_Xong_Nuoc_Khi" )
      S_Coil( "Q_AUTO_V2_Xuc_Khi" )
      R_Coil( "TG_can_Xong_Nuoc_Khi" )
   END_RUNG
   RUNG wire#w1
      Contact( "TG_Can_Xong_CO2" )
      S_Coil( "Q_AUTO_V2_CO2" )
      R_Coil( "TG_Can_Xong_CO2" )
   END_RUNG
   RUNG wire#w1
      Contact( "Q_AUTO_V2_Xuc_Khi" )
      { S7_Templates := "SrcType := Real" } LE_Contact(in1 := "Act_Can_CO2", in2 := 0.0)
      S_Coil( "TG_Can_Xong_CO2" )
      R_Coil( "Q_AUTO_V2_CO2" )
   END_RUNG
   RUNG wire#w1
      Contact( "Q_AUTO_V2_Xuc_Khi" )
      { S7_Templates := "SrcType := Real" } LE_Contact(in1 := "Act_can_nuoc_xuc_khi", in2 := 0.0)
      S_Coil( "TG_can_Xong_Nuoc_Khi" )
      R_Coil( "Q_AUTO_V2_Xuc_Khi" )
   END_RUNG
   RUNG wire#w1
      Contact( "TG_Can_Xong_CO2" )
      Contact( "TG_can_Xong_Nuoc_Khi" )
      R_Coil( "Q_AUTO_LAM_LANH" )
      S_Coil( "Q_AUTO_BOM_2" )
   END_RUNG
   RUNG wire#w1
      Contact( "Q_AUTO_BOM_2" )
      { S7_Templates := "SrcType := Real" } LE_Contact(in1 := "Act_bon_2", in2 := 0.0)
      S_Coil( "TG_Step_3" )
      R_Coil( "TG_Can_Xong_CO2" )
      R_Coil( "TG_can_Xong_Nuoc_Khi" )
      R_Coil( "Q_AUTO_BOM_2" )
      R_Coil( "TG_Step_2" )
   END_RUNG
   // the same network as SCL:
   #_w1 := "TG_Step_2" AND NOT "P6";   // rising edge
   "P6" := "TG_Step_2";
   IF #_w1 THEN "Q_AUTO_LAM_LANH" := TRUE; END_IF;
   IF "TG_Step_2" AND "TG_can_Xong_Nuoc_Khi" THEN
       "Q_AUTO_V2_Xuc_Khi" := TRUE;
       "TG_can_Xong_Nuoc_Khi" := FALSE;
   END_IF;
   IF "TG_Step_2" AND "TG_Can_Xong_CO2" THEN
       "Q_AUTO_V2_CO2" := TRUE;
       "TG_Can_Xong_CO2" := FALSE;
   END_IF;
   IF "TG_Step_2" AND "Q_AUTO_V2_Xuc_Khi" AND ("Act_Can_CO2" <= 0.0) THEN
       "TG_Can_Xong_CO2" := TRUE;
       "Q_AUTO_V2_CO2" := FALSE;
   END_IF;
   IF "TG_Step_2" AND "Q_AUTO_V2_Xuc_Khi" AND ("Act_can_nuoc_xuc_khi" <= 0.0) THEN
       "TG_can_Xong_Nuoc_Khi" := TRUE;
       "Q_AUTO_V2_Xuc_Khi" := FALSE;
   END_IF;
   IF "TG_Step_2" AND "TG_Can_Xong_CO2" AND "TG_can_Xong_Nuoc_Khi" THEN
       "Q_AUTO_LAM_LANH" := FALSE;
       "Q_AUTO_BOM_2" := TRUE;
   END_IF;
   IF "TG_Step_2" AND "Q_AUTO_BOM_2" AND ("Act_bon_2" <= 0.0) THEN
       "TG_Step_3" := TRUE;
       "TG_Can_Xong_CO2" := FALSE;
       "TG_can_Xong_Nuoc_Khi" := FALSE;
   END_IF;
   #_w2 := "TG_Step_2" AND "Q_AUTO_BOM_2" AND ("Act_bon_2" <= 0.0);
   IF #_w2 THEN
       "Q_AUTO_BOM_2" := FALSE;
       "TG_Step_2" := FALSE;
   END_IF;
END_REGION

REGION Network 5
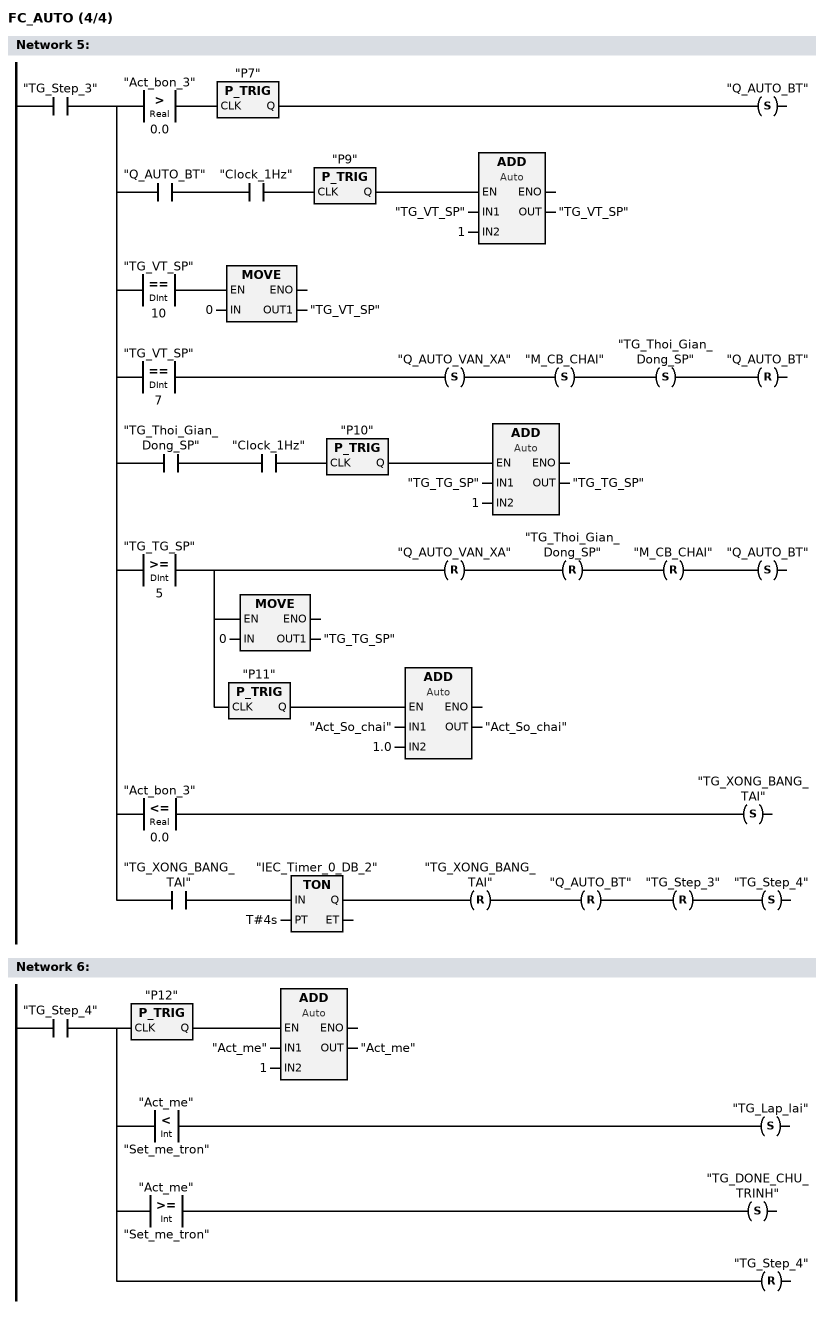
   #_w1 := "TG_Step_3" AND ("Act_bon_3" > 0.0);
   #_w2 := #_w1 AND NOT "P7";   // rising edge
   "P7" := #_w1;
   IF #_w2 THEN "Q_AUTO_BT" := TRUE; END_IF;
   #_w3 := "TG_Step_3" AND "Q_AUTO_BT" AND "Clock_1Hz";
   #_w4 := #_w3 AND NOT "P9";   // rising edge
   "P9" := #_w3;
   IF #_w4 THEN "TG_VT_SP" := "TG_VT_SP" + 1; END_IF;
   IF "TG_Step_3" AND ("TG_VT_SP" = 10) THEN "TG_VT_SP" := 0; END_IF;
   IF "TG_Step_3" AND ("TG_VT_SP" = 7) THEN
       "Q_AUTO_VAN_XA" := TRUE;
       "M_CB_CHAI" := TRUE;
       "TG_Thoi_Gian_Dong_SP" := TRUE;
       "Q_AUTO_BT" := FALSE;
   END_IF;
   #_w5 := "TG_Step_3" AND "TG_Thoi_Gian_Dong_SP" AND "Clock_1Hz";
   #_w6 := #_w5 AND NOT "P10";   // rising edge
   "P10" := #_w5;
   IF #_w6 THEN "TG_TG_SP" := "TG_TG_SP" + 1; END_IF;
   #_w7 := "TG_Step_3" AND ("TG_TG_SP" >= 5);
   IF #_w7 THEN
       "Q_AUTO_VAN_XA" := FALSE;
       "TG_Thoi_Gian_Dong_SP" := FALSE;
       "M_CB_CHAI" := FALSE;
       "Q_AUTO_BT" := TRUE;
       "TG_TG_SP" := 0;
   END_IF;
   #_w8 := #_w7 AND NOT "P11";   // rising edge
   "P11" := #_w7;
   IF #_w8 THEN "Act_So_chai" := "Act_So_chai" + 1.0; END_IF;
   IF "TG_Step_3" AND ("Act_bon_3" <= 0.0) THEN "TG_XONG_BANG_TAI" := TRUE; END_IF;
   "IEC_Timer_0_DB_2".TON(IN := "TG_Step_3" AND "TG_XONG_BANG_TAI", PT := T#4s);
   IF "IEC_Timer_0_DB_2".Q THEN
       "TG_XONG_BANG_TAI" := FALSE;
       "Q_AUTO_BT" := FALSE;
       "TG_Step_3" := FALSE;
       "TG_Step_4" := TRUE;
   END_IF;
END_REGION

REGION Network 6
   RUNG wire#powerrail
      Contact( "TG_Step_4" )
      wire#w1
      P_Trig( "P12" )
      Add(in1 := "Act_me", in2 := 1, out => "Act_me")
   END_RUNG
   RUNG wire#w1
      { S7_Templates := "SrcType := Int" } LT_Contact(in1 := "Act_me", in2 := "Set_me_tron")
      S_Coil( "TG_Lap_lai" )
   END_RUNG
   RUNG wire#w1
      { S7_Templates := "SrcType := Int" } GE_Contact(in1 := "Act_me", in2 := "Set_me_tron")
      S_Coil( "TG_DONE_CHU_TRINH" )
   END_RUNG
   RUNG wire#w1
      R_Coil( "TG_Step_4" )
   END_RUNG
   // the same network as SCL:
   #_w1 := "TG_Step_4" AND NOT "P12";   // rising edge
   "P12" := "TG_Step_4";
   IF #_w1 THEN "Act_me" := "Act_me" + 1; END_IF;
   IF "TG_Step_4" AND ("Act_me" < "Set_me_tron") THEN "TG_Lap_lai" := TRUE; END_IF;
   IF "TG_Step_4" AND ("Act_me" >= "Set_me_tron") THEN "TG_DONE_CHU_TRINH" := TRUE; END_IF;
   IF "TG_Step_4" THEN "TG_Step_4" := FALSE; END_IF;
END_REGION
END_FUNCTION

FUNCTION "FC_MANUAL" : Void   // FC3, LAD
{ S7_Optimized_Access := 'TRUE' }
VERSION : 0.1
BEGIN

REGION Network 1: Bom_1
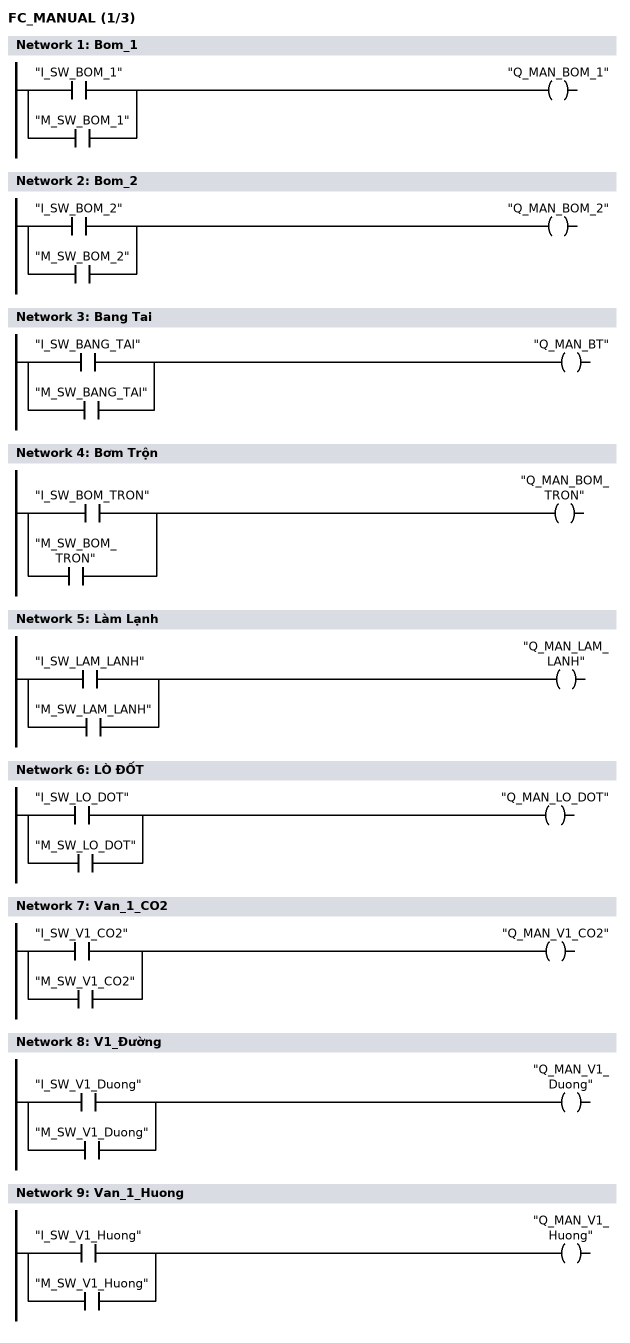
   RUNG wire#powerrail
      Contact( "I_SW_BOM_1" )
      wire#w1
      Coil( "Q_MAN_BOM_1" )
   END_RUNG
   RUNG wire#powerrail
      Contact( "M_SW_BOM_1" )
   END_RUNG wire#w1
   // the same network as SCL:
   "Q_MAN_BOM_1" := "I_SW_BOM_1" OR "M_SW_BOM_1";
END_REGION

REGION Network 2: Bom_2
   RUNG wire#powerrail
      Contact( "I_SW_BOM_2" )
      wire#w1
      Coil( "Q_MAN_BOM_2" )
   END_RUNG
   RUNG wire#powerrail
      Contact( "M_SW_BOM_2" )
   END_RUNG wire#w1
   // the same network as SCL:
   "Q_MAN_BOM_2" := "I_SW_BOM_2" OR "M_SW_BOM_2";
END_REGION

REGION Network 3: Bang Tai
   RUNG wire#powerrail
      Contact( "I_SW_BANG_TAI" )
      wire#w1
      Coil( "Q_MAN_BT" )
   END_RUNG
   RUNG wire#powerrail
      Contact( "M_SW_BANG_TAI" )
   END_RUNG wire#w1
   // the same network as SCL:
   "Q_MAN_BT" := "I_SW_BANG_TAI" OR "M_SW_BANG_TAI";
END_REGION

REGION Network 4: Bơm Trộn
   RUNG wire#powerrail
      Contact( "I_SW_BOM_TRON" )
      wire#w1
      Coil( "Q_MAN_BOM_TRON" )
   END_RUNG
   RUNG wire#powerrail
      Contact( "M_SW_BOM_TRON" )
   END_RUNG wire#w1
   // the same network as SCL:
   "Q_MAN_BOM_TRON" := "I_SW_BOM_TRON" OR "M_SW_BOM_TRON";
END_REGION

REGION Network 5: Làm Lạnh
   RUNG wire#powerrail
      Contact( "I_SW_LAM_LANH" )
      wire#w1
      Coil( "Q_MAN_LAM_LANH" )
   END_RUNG
   RUNG wire#powerrail
      Contact( "M_SW_LAM_LANH" )
   END_RUNG wire#w1
   // the same network as SCL:
   "Q_MAN_LAM_LANH" := "I_SW_LAM_LANH" OR "M_SW_LAM_LANH";
END_REGION

REGION Network 6: LÒ ĐỐT
   RUNG wire#powerrail
      Contact( "I_SW_LO_DOT" )
      wire#w1
      Coil( "Q_MAN_LO_DOT" )
   END_RUNG
   RUNG wire#powerrail
      Contact( "M_SW_LO_DOT" )
   END_RUNG wire#w1
   // the same network as SCL:
   "Q_MAN_LO_DOT" := "I_SW_LO_DOT" OR "M_SW_LO_DOT";
END_REGION

REGION Network 7: Van_1_CO2
   RUNG wire#powerrail
      Contact( "I_SW_V1_CO2" )
      wire#w1
      Coil( "Q_MAN_V1_CO2" )
   END_RUNG
   RUNG wire#powerrail
      Contact( "M_SW_V1_CO2" )
   END_RUNG wire#w1
   // the same network as SCL:
   "Q_MAN_V1_CO2" := "I_SW_V1_CO2" OR "M_SW_V1_CO2";
END_REGION

REGION Network 8: V1_Đường
   RUNG wire#powerrail
      Contact( "I_SW_V1_Duong" )
      wire#w1
      Coil( "Q_MAN_V1_Duong" )
   END_RUNG
   RUNG wire#powerrail
      Contact( "M_SW_V1_Duong" )
   END_RUNG wire#w1
   // the same network as SCL:
   "Q_MAN_V1_Duong" := "I_SW_V1_Duong" OR "M_SW_V1_Duong";
END_REGION

REGION Network 9: Van_1_Huong
   RUNG wire#powerrail
      Contact( "I_SW_V1_Huong" )
      wire#w1
      Coil( "Q_MAN_V1_Huong" )
   END_RUNG
   RUNG wire#powerrail
      Contact( "M_SW_V1_Huong" )
   END_RUNG wire#w1
   // the same network as SCL:
   "Q_MAN_V1_Huong" := "I_SW_V1_Huong" OR "M_SW_V1_Huong";
END_REGION

REGION Network 10: Van_1_Màu
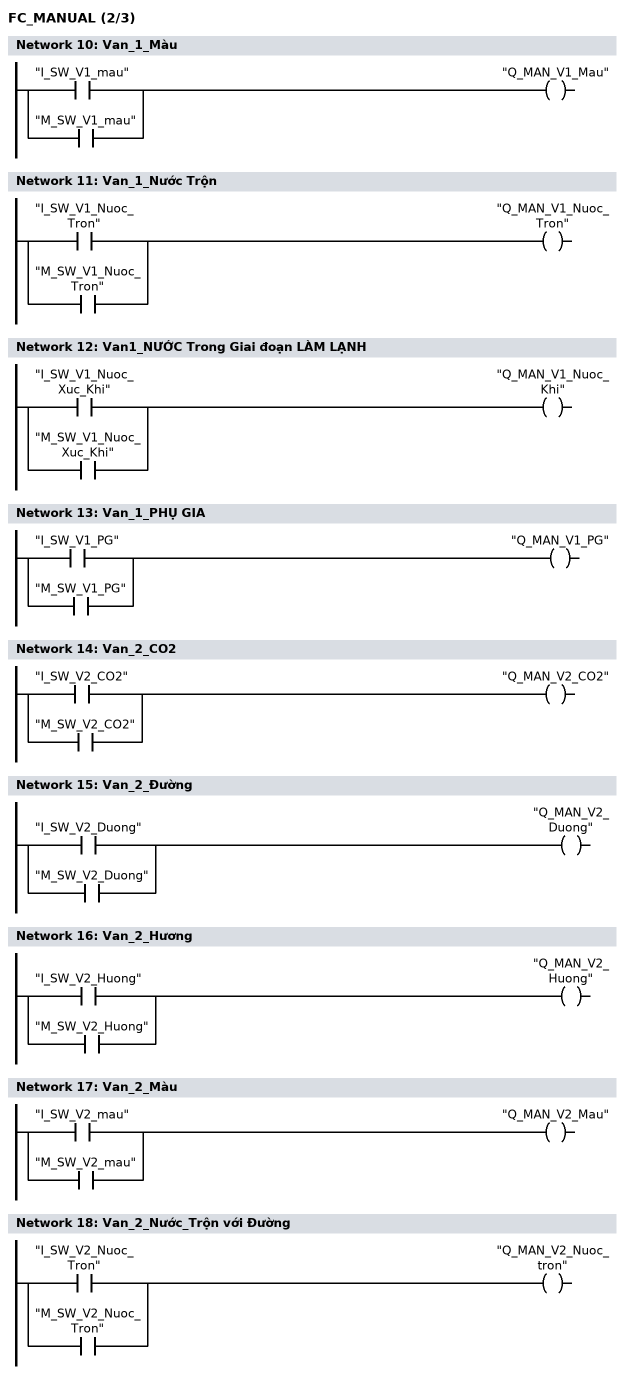
   RUNG wire#powerrail
      Contact( "I_SW_V1_mau" )
      wire#w1
      Coil( "Q_MAN_V1_Mau" )
   END_RUNG
   RUNG wire#powerrail
      Contact( "M_SW_V1_mau" )
   END_RUNG wire#w1
   // the same network as SCL:
   "Q_MAN_V1_Mau" := "I_SW_V1_mau" OR "M_SW_V1_mau";
END_REGION

REGION Network 11: Van_1_Nước Trộn
   RUNG wire#powerrail
      Contact( "I_SW_V1_Nuoc_Tron" )
      wire#w1
      Coil( "Q_MAN_V1_Nuoc_Tron" )
   END_RUNG
   RUNG wire#powerrail
      Contact( "M_SW_V1_Nuoc_Tron" )
   END_RUNG wire#w1
   // the same network as SCL:
   "Q_MAN_V1_Nuoc_Tron" := "I_SW_V1_Nuoc_Tron" OR "M_SW_V1_Nuoc_Tron";
END_REGION

REGION Network 12: Van1_NƯỚC Trong Giai đoạn LÀM LẠNH
   RUNG wire#powerrail
      Contact( "I_SW_V1_Nuoc_Xuc_Khi" )
      wire#w1
      Coil( "Q_MAN_V1_Nuoc_Khi" )
   END_RUNG
   RUNG wire#powerrail
      Contact( "M_SW_V1_Nuoc_Xuc_Khi" )
   END_RUNG wire#w1
   // the same network as SCL:
   "Q_MAN_V1_Nuoc_Khi" := "I_SW_V1_Nuoc_Xuc_Khi" OR "M_SW_V1_Nuoc_Xuc_Khi";
END_REGION

REGION Network 13: Van_1_PHỤ GIA
   RUNG wire#powerrail
      Contact( "I_SW_V1_PG" )
      wire#w1
      Coil( "Q_MAN_V1_PG" )
   END_RUNG
   RUNG wire#powerrail
      Contact( "M_SW_V1_PG" )
   END_RUNG wire#w1
   // the same network as SCL:
   "Q_MAN_V1_PG" := "I_SW_V1_PG" OR "M_SW_V1_PG";
END_REGION

REGION Network 14: Van_2_CO2
   RUNG wire#powerrail
      Contact( "I_SW_V2_CO2" )
      wire#w1
      Coil( "Q_MAN_V2_CO2" )
   END_RUNG
   RUNG wire#powerrail
      Contact( "M_SW_V2_CO2" )
   END_RUNG wire#w1
   // the same network as SCL:
   "Q_MAN_V2_CO2" := "I_SW_V2_CO2" OR "M_SW_V2_CO2";
END_REGION

REGION Network 15: Van_2_Đường
   RUNG wire#powerrail
      Contact( "I_SW_V2_Duong" )
      wire#w1
      Coil( "Q_MAN_V2_Duong" )
   END_RUNG
   RUNG wire#powerrail
      Contact( "M_SW_V2_Duong" )
   END_RUNG wire#w1
   // the same network as SCL:
   "Q_MAN_V2_Duong" := "I_SW_V2_Duong" OR "M_SW_V2_Duong";
END_REGION

REGION Network 16: Van_2_Hương
   RUNG wire#powerrail
      Contact( "I_SW_V2_Huong" )
      wire#w1
      Coil( "Q_MAN_V2_Huong" )
   END_RUNG
   RUNG wire#powerrail
      Contact( "M_SW_V2_Huong" )
   END_RUNG wire#w1
   // the same network as SCL:
   "Q_MAN_V2_Huong" := "I_SW_V2_Huong" OR "M_SW_V2_Huong";
END_REGION

REGION Network 17: Van_2_Màu
   RUNG wire#powerrail
      Contact( "I_SW_V2_mau" )
      wire#w1
      Coil( "Q_MAN_V2_Mau" )
   END_RUNG
   RUNG wire#powerrail
      Contact( "M_SW_V2_mau" )
   END_RUNG wire#w1
   // the same network as SCL:
   "Q_MAN_V2_Mau" := "I_SW_V2_mau" OR "M_SW_V2_mau";
END_REGION

REGION Network 18: Van_2_Nước_Trộn với Đường
   RUNG wire#powerrail
      Contact( "I_SW_V2_Nuoc_Tron" )
      wire#w1
      Coil( "Q_MAN_V2_Nuoc_tron" )
   END_RUNG
   RUNG wire#powerrail
      Contact( "M_SW_V2_Nuoc_Tron" )
   END_RUNG wire#w1
   // the same network as SCL:
   "Q_MAN_V2_Nuoc_tron" := "I_SW_V2_Nuoc_Tron" OR "M_SW_V2_Nuoc_Tron";
END_REGION

REGION Network 19: Van_2_ NƯớc LÀm lạnh
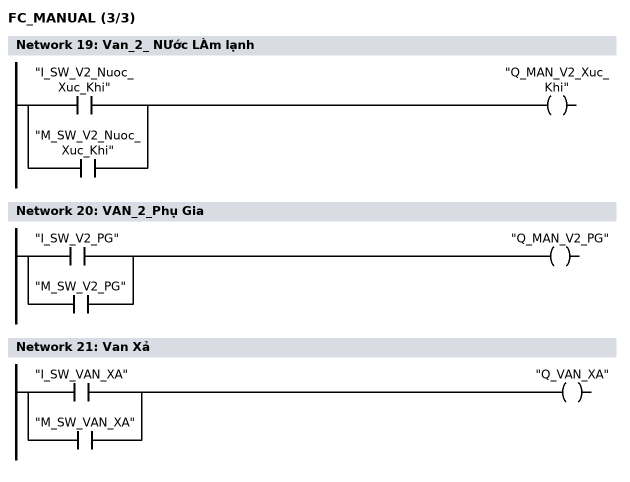
   RUNG wire#powerrail
      Contact( "I_SW_V2_Nuoc_Xuc_Khi" )
      wire#w1
      Coil( "Q_MAN_V2_Xuc_Khi" )
   END_RUNG
   RUNG wire#powerrail
      Contact( "M_SW_V2_Nuoc_Xuc_Khi" )
   END_RUNG wire#w1
   // the same network as SCL:
   "Q_MAN_V2_Xuc_Khi" := "I_SW_V2_Nuoc_Xuc_Khi" OR "M_SW_V2_Nuoc_Xuc_Khi";
END_REGION

REGION Network 20: VAN_2_Phụ Gia
   RUNG wire#powerrail
      Contact( "I_SW_V2_PG" )
      wire#w1
      Coil( "Q_MAN_V2_PG" )
   END_RUNG
   RUNG wire#powerrail
      Contact( "M_SW_V2_PG" )
   END_RUNG wire#w1
   // the same network as SCL:
   "Q_MAN_V2_PG" := "I_SW_V2_PG" OR "M_SW_V2_PG";
END_REGION

REGION Network 21: Van Xả
   RUNG wire#powerrail
      Contact( "I_SW_VAN_XA" )
      wire#w1
      Coil( "Q_VAN_XA" )
   END_RUNG
   RUNG wire#powerrail
      Contact( "M_SW_VAN_XA" )
   END_RUNG wire#w1
   // the same network as SCL:
   "Q_VAN_XA" := "I_SW_VAN_XA" OR "M_SW_VAN_XA";
END_REGION
END_FUNCTION

FUNCTION "FC_OUTPUT" : Void   // FC4, LAD
{ S7_Optimized_Access := 'TRUE' }
VERSION : 0.1
BEGIN

REGION Network 1
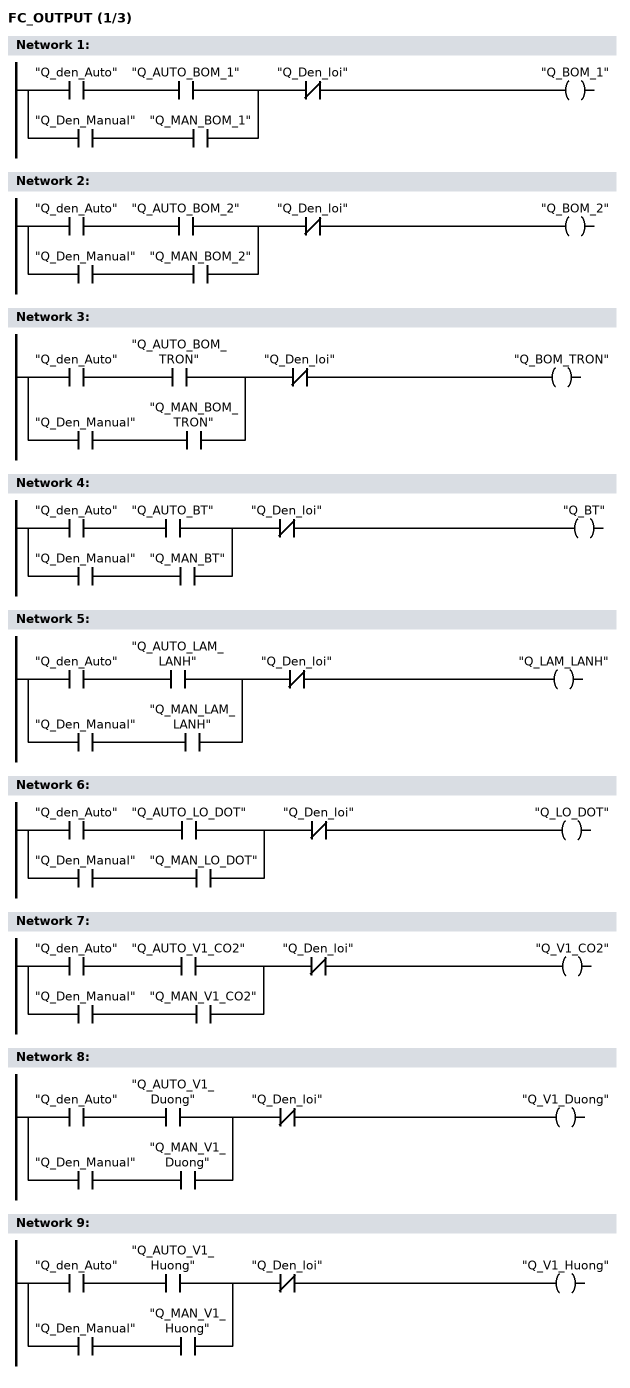
   RUNG wire#powerrail
      Contact( "Q_den_Auto" )
      Contact( "Q_AUTO_BOM_1" )
      wire#w1
      I_Contact( "Q_Den_loi" )
      Coil( "Q_BOM_1" )
   END_RUNG
   RUNG wire#powerrail
      Contact( "Q_Den_Manual" )
      Contact( "Q_MAN_BOM_1" )
   END_RUNG wire#w1
   // the same network as SCL:
   "Q_BOM_1" := (("Q_den_Auto" AND "Q_AUTO_BOM_1") OR ("Q_Den_Manual" AND "Q_MAN_BOM_1")) AND NOT "Q_Den_loi";
END_REGION

REGION Network 2
   RUNG wire#powerrail
      Contact( "Q_den_Auto" )
      Contact( "Q_AUTO_BOM_2" )
      wire#w1
      I_Contact( "Q_Den_loi" )
      Coil( "Q_BOM_2" )
   END_RUNG
   RUNG wire#powerrail
      Contact( "Q_Den_Manual" )
      Contact( "Q_MAN_BOM_2" )
   END_RUNG wire#w1
   // the same network as SCL:
   "Q_BOM_2" := (("Q_den_Auto" AND "Q_AUTO_BOM_2") OR ("Q_Den_Manual" AND "Q_MAN_BOM_2")) AND NOT "Q_Den_loi";
END_REGION

REGION Network 3
   RUNG wire#powerrail
      Contact( "Q_den_Auto" )
      Contact( "Q_AUTO_BOM_TRON" )
      wire#w1
      I_Contact( "Q_Den_loi" )
      Coil( "Q_BOM_TRON" )
   END_RUNG
   RUNG wire#powerrail
      Contact( "Q_Den_Manual" )
      Contact( "Q_MAN_BOM_TRON" )
   END_RUNG wire#w1
   // the same network as SCL:
   "Q_BOM_TRON" := (("Q_den_Auto" AND "Q_AUTO_BOM_TRON") OR ("Q_Den_Manual" AND "Q_MAN_BOM_TRON")) AND NOT "Q_Den_loi";
END_REGION

REGION Network 4
   RUNG wire#powerrail
      Contact( "Q_den_Auto" )
      Contact( "Q_AUTO_BT" )
      wire#w1
      I_Contact( "Q_Den_loi" )
      Coil( "Q_BT" )
   END_RUNG
   RUNG wire#powerrail
      Contact( "Q_Den_Manual" )
      Contact( "Q_MAN_BT" )
   END_RUNG wire#w1
   // the same network as SCL:
   "Q_BT" := (("Q_den_Auto" AND "Q_AUTO_BT") OR ("Q_Den_Manual" AND "Q_MAN_BT")) AND NOT "Q_Den_loi";
END_REGION

REGION Network 5
   RUNG wire#powerrail
      Contact( "Q_den_Auto" )
      Contact( "Q_AUTO_LAM_LANH" )
      wire#w1
      I_Contact( "Q_Den_loi" )
      Coil( "Q_LAM_LANH" )
   END_RUNG
   RUNG wire#powerrail
      Contact( "Q_Den_Manual" )
      Contact( "Q_MAN_LAM_LANH" )
   END_RUNG wire#w1
   // the same network as SCL:
   "Q_LAM_LANH" := (("Q_den_Auto" AND "Q_AUTO_LAM_LANH") OR ("Q_Den_Manual" AND "Q_MAN_LAM_LANH")) AND NOT "Q_Den_loi";
END_REGION

REGION Network 6
   RUNG wire#powerrail
      Contact( "Q_den_Auto" )
      Contact( "Q_AUTO_LO_DOT" )
      wire#w1
      I_Contact( "Q_Den_loi" )
      Coil( "Q_LO_DOT" )
   END_RUNG
   RUNG wire#powerrail
      Contact( "Q_Den_Manual" )
      Contact( "Q_MAN_LO_DOT" )
   END_RUNG wire#w1
   // the same network as SCL:
   "Q_LO_DOT" := (("Q_den_Auto" AND "Q_AUTO_LO_DOT") OR ("Q_Den_Manual" AND "Q_MAN_LO_DOT")) AND NOT "Q_Den_loi";
END_REGION

REGION Network 7
   RUNG wire#powerrail
      Contact( "Q_den_Auto" )
      Contact( "Q_AUTO_V1_CO2" )
      wire#w1
      I_Contact( "Q_Den_loi" )
      Coil( "Q_V1_CO2" )
   END_RUNG
   RUNG wire#powerrail
      Contact( "Q_Den_Manual" )
      Contact( "Q_MAN_V1_CO2" )
   END_RUNG wire#w1
   // the same network as SCL:
   "Q_V1_CO2" := (("Q_den_Auto" AND "Q_AUTO_V1_CO2") OR ("Q_Den_Manual" AND "Q_MAN_V1_CO2")) AND NOT "Q_Den_loi";
END_REGION

REGION Network 8
   RUNG wire#powerrail
      Contact( "Q_den_Auto" )
      Contact( "Q_AUTO_V1_Duong" )
      wire#w1
      I_Contact( "Q_Den_loi" )
      Coil( "Q_V1_Duong" )
   END_RUNG
   RUNG wire#powerrail
      Contact( "Q_Den_Manual" )
      Contact( "Q_MAN_V1_Duong" )
   END_RUNG wire#w1
   // the same network as SCL:
   "Q_V1_Duong" := (("Q_den_Auto" AND "Q_AUTO_V1_Duong") OR ("Q_Den_Manual" AND "Q_MAN_V1_Duong")) AND NOT "Q_Den_loi";
END_REGION

REGION Network 9
   RUNG wire#powerrail
      Contact( "Q_den_Auto" )
      Contact( "Q_AUTO_V1_Huong" )
      wire#w1
      I_Contact( "Q_Den_loi" )
      Coil( "Q_V1_Huong" )
   END_RUNG
   RUNG wire#powerrail
      Contact( "Q_Den_Manual" )
      Contact( "Q_MAN_V1_Huong" )
   END_RUNG wire#w1
   // the same network as SCL:
   "Q_V1_Huong" := (("Q_den_Auto" AND "Q_AUTO_V1_Huong") OR ("Q_Den_Manual" AND "Q_MAN_V1_Huong")) AND NOT "Q_Den_loi";
END_REGION

REGION Network 10
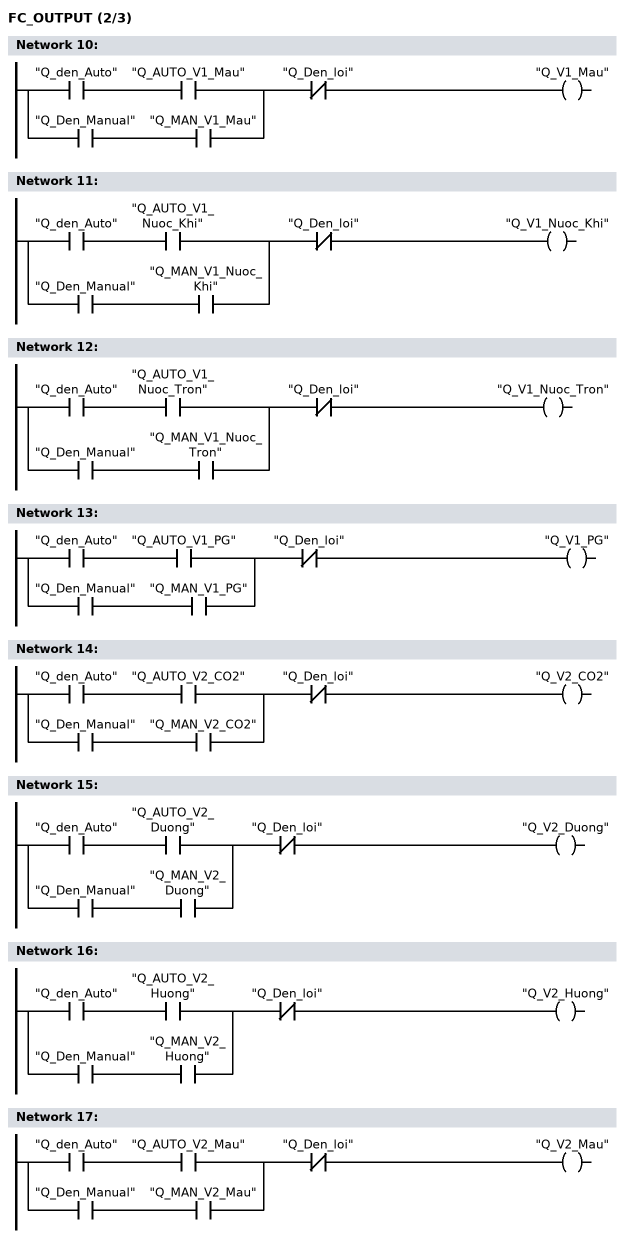
   RUNG wire#powerrail
      Contact( "Q_den_Auto" )
      Contact( "Q_AUTO_V1_Mau" )
      wire#w1
      I_Contact( "Q_Den_loi" )
      Coil( "Q_V1_Mau" )
   END_RUNG
   RUNG wire#powerrail
      Contact( "Q_Den_Manual" )
      Contact( "Q_MAN_V1_Mau" )
   END_RUNG wire#w1
   // the same network as SCL:
   "Q_V1_Mau" := (("Q_den_Auto" AND "Q_AUTO_V1_Mau") OR ("Q_Den_Manual" AND "Q_MAN_V1_Mau")) AND NOT "Q_Den_loi";
END_REGION

REGION Network 11
   RUNG wire#powerrail
      Contact( "Q_den_Auto" )
      Contact( "Q_AUTO_V1_Nuoc_Khi" )
      wire#w1
      I_Contact( "Q_Den_loi" )
      Coil( "Q_V1_Nuoc_Khi" )
   END_RUNG
   RUNG wire#powerrail
      Contact( "Q_Den_Manual" )
      Contact( "Q_MAN_V1_Nuoc_Khi" )
   END_RUNG wire#w1
   // the same network as SCL:
   "Q_V1_Nuoc_Khi" := (("Q_den_Auto" AND "Q_AUTO_V1_Nuoc_Khi") OR ("Q_Den_Manual" AND "Q_MAN_V1_Nuoc_Khi")) AND NOT "Q_Den_loi";
END_REGION

REGION Network 12
   RUNG wire#powerrail
      Contact( "Q_den_Auto" )
      Contact( "Q_AUTO_V1_Nuoc_Tron" )
      wire#w1
      I_Contact( "Q_Den_loi" )
      Coil( "Q_V1_Nuoc_Tron" )
   END_RUNG
   RUNG wire#powerrail
      Contact( "Q_Den_Manual" )
      Contact( "Q_MAN_V1_Nuoc_Tron" )
   END_RUNG wire#w1
   // the same network as SCL:
   "Q_V1_Nuoc_Tron" := (("Q_den_Auto" AND "Q_AUTO_V1_Nuoc_Tron") OR ("Q_Den_Manual" AND "Q_MAN_V1_Nuoc_Tron")) AND NOT "Q_Den_loi";
END_REGION

REGION Network 13
   RUNG wire#powerrail
      Contact( "Q_den_Auto" )
      Contact( "Q_AUTO_V1_PG" )
      wire#w1
      I_Contact( "Q_Den_loi" )
      Coil( "Q_V1_PG" )
   END_RUNG
   RUNG wire#powerrail
      Contact( "Q_Den_Manual" )
      Contact( "Q_MAN_V1_PG" )
   END_RUNG wire#w1
   // the same network as SCL:
   "Q_V1_PG" := (("Q_den_Auto" AND "Q_AUTO_V1_PG") OR ("Q_Den_Manual" AND "Q_MAN_V1_PG")) AND NOT "Q_Den_loi";
END_REGION

REGION Network 14
   RUNG wire#powerrail
      Contact( "Q_den_Auto" )
      Contact( "Q_AUTO_V2_CO2" )
      wire#w1
      I_Contact( "Q_Den_loi" )
      Coil( "Q_V2_CO2" )
   END_RUNG
   RUNG wire#powerrail
      Contact( "Q_Den_Manual" )
      Contact( "Q_MAN_V2_CO2" )
   END_RUNG wire#w1
   // the same network as SCL:
   "Q_V2_CO2" := (("Q_den_Auto" AND "Q_AUTO_V2_CO2") OR ("Q_Den_Manual" AND "Q_MAN_V2_CO2")) AND NOT "Q_Den_loi";
END_REGION

REGION Network 15
   RUNG wire#powerrail
      Contact( "Q_den_Auto" )
      Contact( "Q_AUTO_V2_Duong" )
      wire#w1
      I_Contact( "Q_Den_loi" )
      Coil( "Q_V2_Duong" )
   END_RUNG
   RUNG wire#powerrail
      Contact( "Q_Den_Manual" )
      Contact( "Q_MAN_V2_Duong" )
   END_RUNG wire#w1
   // the same network as SCL:
   "Q_V2_Duong" := (("Q_den_Auto" AND "Q_AUTO_V2_Duong") OR ("Q_Den_Manual" AND "Q_MAN_V2_Duong")) AND NOT "Q_Den_loi";
END_REGION

REGION Network 16
   RUNG wire#powerrail
      Contact( "Q_den_Auto" )
      Contact( "Q_AUTO_V2_Huong" )
      wire#w1
      I_Contact( "Q_Den_loi" )
      Coil( "Q_V2_Huong" )
   END_RUNG
   RUNG wire#powerrail
      Contact( "Q_Den_Manual" )
      Contact( "Q_MAN_V2_Huong" )
   END_RUNG wire#w1
   // the same network as SCL:
   "Q_V2_Huong" := (("Q_den_Auto" AND "Q_AUTO_V2_Huong") OR ("Q_Den_Manual" AND "Q_MAN_V2_Huong")) AND NOT "Q_Den_loi";
END_REGION

REGION Network 17
   RUNG wire#powerrail
      Contact( "Q_den_Auto" )
      Contact( "Q_AUTO_V2_Mau" )
      wire#w1
      I_Contact( "Q_Den_loi" )
      Coil( "Q_V2_Mau" )
   END_RUNG
   RUNG wire#powerrail
      Contact( "Q_Den_Manual" )
      Contact( "Q_MAN_V2_Mau" )
   END_RUNG wire#w1
   // the same network as SCL:
   "Q_V2_Mau" := (("Q_den_Auto" AND "Q_AUTO_V2_Mau") OR ("Q_Den_Manual" AND "Q_MAN_V2_Mau")) AND NOT "Q_Den_loi";
END_REGION

REGION Network 18
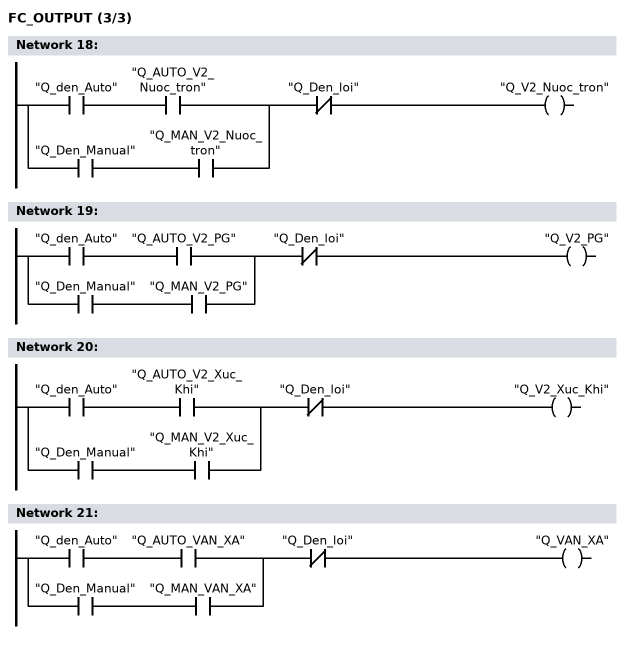
   RUNG wire#powerrail
      Contact( "Q_den_Auto" )
      Contact( "Q_AUTO_V2_Nuoc_tron" )
      wire#w1
      I_Contact( "Q_Den_loi" )
      Coil( "Q_V2_Nuoc_tron" )
   END_RUNG
   RUNG wire#powerrail
      Contact( "Q_Den_Manual" )
      Contact( "Q_MAN_V2_Nuoc_tron" )
   END_RUNG wire#w1
   // the same network as SCL:
   "Q_V2_Nuoc_tron" := (("Q_den_Auto" AND "Q_AUTO_V2_Nuoc_tron") OR ("Q_Den_Manual" AND "Q_MAN_V2_Nuoc_tron")) AND NOT "Q_Den_loi";
END_REGION

REGION Network 19
   RUNG wire#powerrail
      Contact( "Q_den_Auto" )
      Contact( "Q_AUTO_V2_PG" )
      wire#w1
      I_Contact( "Q_Den_loi" )
      Coil( "Q_V2_PG" )
   END_RUNG
   RUNG wire#powerrail
      Contact( "Q_Den_Manual" )
      Contact( "Q_MAN_V2_PG" )
   END_RUNG wire#w1
   // the same network as SCL:
   "Q_V2_PG" := (("Q_den_Auto" AND "Q_AUTO_V2_PG") OR ("Q_Den_Manual" AND "Q_MAN_V2_PG")) AND NOT "Q_Den_loi";
END_REGION

REGION Network 20
   RUNG wire#powerrail
      Contact( "Q_den_Auto" )
      Contact( "Q_AUTO_V2_Xuc_Khi" )
      wire#w1
      I_Contact( "Q_Den_loi" )
      Coil( "Q_V2_Xuc_Khi" )
   END_RUNG
   RUNG wire#powerrail
      Contact( "Q_Den_Manual" )
      Contact( "Q_MAN_V2_Xuc_Khi" )
   END_RUNG wire#w1
   // the same network as SCL:
   "Q_V2_Xuc_Khi" := (("Q_den_Auto" AND "Q_AUTO_V2_Xuc_Khi") OR ("Q_Den_Manual" AND "Q_MAN_V2_Xuc_Khi")) AND NOT "Q_Den_loi";
END_REGION

REGION Network 21
   RUNG wire#powerrail
      Contact( "Q_den_Auto" )
      Contact( "Q_AUTO_VAN_XA" )
      wire#w1
      I_Contact( "Q_Den_loi" )
      Coil( "Q_VAN_XA" )
   END_RUNG
   RUNG wire#powerrail
      Contact( "Q_Den_Manual" )
      Contact( "Q_MAN_VAN_XA" )
   END_RUNG wire#w1
   // the same network as SCL:
   "Q_VAN_XA" := (("Q_den_Auto" AND "Q_AUTO_VAN_XA") OR ("Q_Den_Manual" AND "Q_MAN_VAN_XA")) AND NOT "Q_Den_loi";
END_REGION
END_FUNCTION

FUNCTION "FC_SIMULATION" : Void   // FC5, LAD
{ S7_Optimized_Access := 'TRUE' }
VERSION : 0.1
   VAR_TEMP   // added for the SCL form of the ladder/FBD networks
      _w1 : Bool;
   END_VAR
BEGIN

REGION Network 1
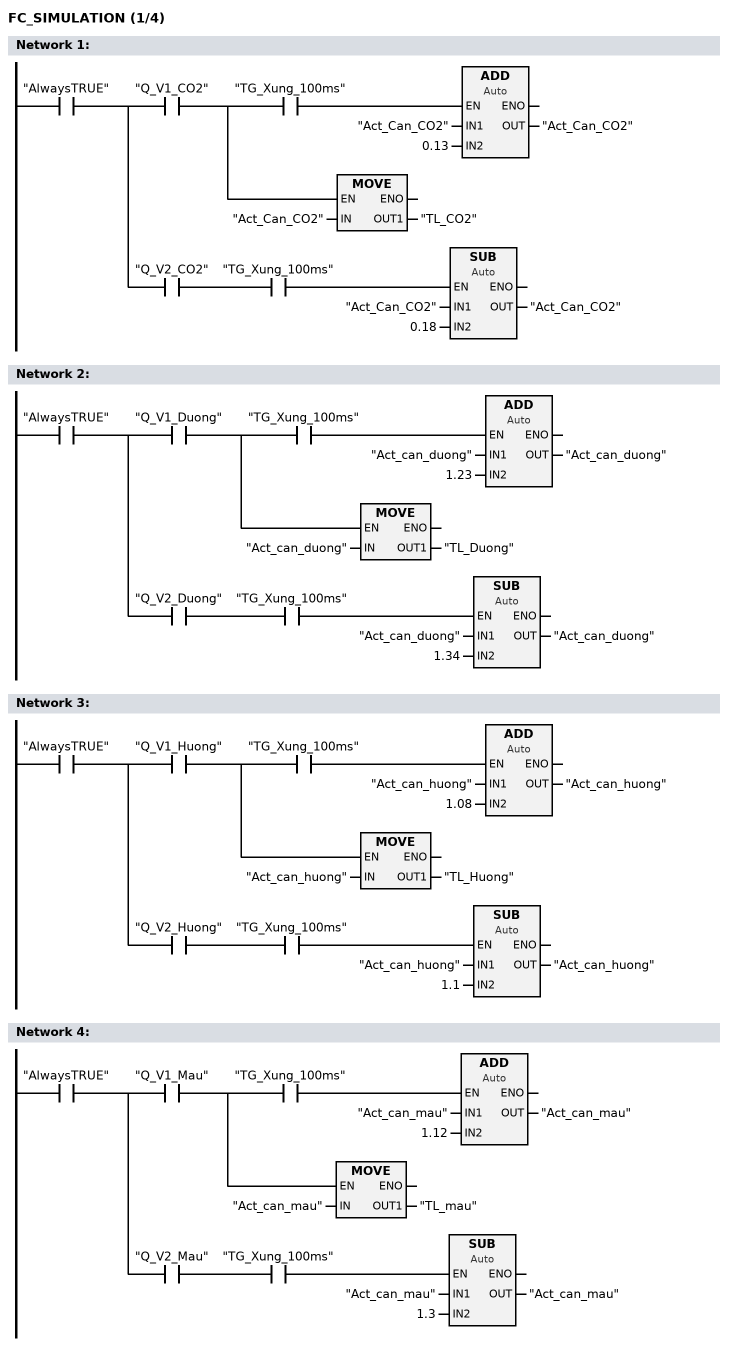
   RUNG wire#powerrail
      Contact( "AlwaysTRUE" )
      wire#w1
      Contact( "Q_V1_CO2" )
      wire#w2
      Contact( "TG_Xung_100ms" )
      Add(in1 := "Act_Can_CO2", in2 := 0.13, out => "Act_Can_CO2")
   END_RUNG
   RUNG wire#w2
      Move(in := "Act_Can_CO2", out1 => "TL_CO2")
   END_RUNG
   RUNG wire#w1
      Contact( "Q_V2_CO2" )
      Contact( "TG_Xung_100ms" )
      Sub(in1 := "Act_Can_CO2", in2 := 0.18, out => "Act_Can_CO2")
   END_RUNG
   // the same network as SCL:
   #_w1 := "AlwaysTRUE" AND "Q_V1_CO2";
   IF #_w1 AND "TG_Xung_100ms" THEN "Act_Can_CO2" := "Act_Can_CO2" + 0.13; END_IF;
   IF #_w1 THEN "TL_CO2" := "Act_Can_CO2"; END_IF;
   IF "AlwaysTRUE" AND "Q_V2_CO2" AND "TG_Xung_100ms" THEN "Act_Can_CO2" := "Act_Can_CO2" - 0.18; END_IF;
END_REGION

REGION Network 2
   RUNG wire#powerrail
      Contact( "AlwaysTRUE" )
      wire#w1
      Contact( "Q_V1_Duong" )
      wire#w2
      Contact( "TG_Xung_100ms" )
      Add(in1 := "Act_can_duong", in2 := 1.23, out => "Act_can_duong")
   END_RUNG
   RUNG wire#w2
      Move(in := "Act_can_duong", out1 => "TL_Duong")
   END_RUNG
   RUNG wire#w1
      Contact( "Q_V2_Duong" )
      Contact( "TG_Xung_100ms" )
      Sub(in1 := "Act_can_duong", in2 := 1.34, out => "Act_can_duong")
   END_RUNG
   // the same network as SCL:
   #_w1 := "AlwaysTRUE" AND "Q_V1_Duong";
   IF #_w1 AND "TG_Xung_100ms" THEN "Act_can_duong" := "Act_can_duong" + 1.23; END_IF;
   IF #_w1 THEN "TL_Duong" := "Act_can_duong"; END_IF;
   IF "AlwaysTRUE" AND "Q_V2_Duong" AND "TG_Xung_100ms" THEN
       "Act_can_duong" := "Act_can_duong" - 1.34;
   END_IF;
END_REGION

REGION Network 3
   RUNG wire#powerrail
      Contact( "AlwaysTRUE" )
      wire#w1
      Contact( "Q_V1_Huong" )
      wire#w2
      Contact( "TG_Xung_100ms" )
      Add(in1 := "Act_can_huong", in2 := 1.08, out => "Act_can_huong")
   END_RUNG
   RUNG wire#w2
      Move(in := "Act_can_huong", out1 => "TL_Huong")
   END_RUNG
   RUNG wire#w1
      Contact( "Q_V2_Huong" )
      Contact( "TG_Xung_100ms" )
      Sub(in1 := "Act_can_huong", in2 := 1.1, out => "Act_can_huong")
   END_RUNG
   // the same network as SCL:
   #_w1 := "AlwaysTRUE" AND "Q_V1_Huong";
   IF #_w1 AND "TG_Xung_100ms" THEN "Act_can_huong" := "Act_can_huong" + 1.08; END_IF;
   IF #_w1 THEN "TL_Huong" := "Act_can_huong"; END_IF;
   IF "AlwaysTRUE" AND "Q_V2_Huong" AND "TG_Xung_100ms" THEN
       "Act_can_huong" := "Act_can_huong" - 1.1;
   END_IF;
END_REGION

REGION Network 4
   RUNG wire#powerrail
      Contact( "AlwaysTRUE" )
      wire#w1
      Contact( "Q_V1_Mau" )
      wire#w2
      Contact( "TG_Xung_100ms" )
      Add(in1 := "Act_can_mau", in2 := 1.12, out => "Act_can_mau")
   END_RUNG
   RUNG wire#w2
      Move(in := "Act_can_mau", out1 => "TL_mau")
   END_RUNG
   RUNG wire#w1
      Contact( "Q_V2_Mau" )
      Contact( "TG_Xung_100ms" )
      Sub(in1 := "Act_can_mau", in2 := 1.3, out => "Act_can_mau")
   END_RUNG
   // the same network as SCL:
   #_w1 := "AlwaysTRUE" AND "Q_V1_Mau";
   IF #_w1 AND "TG_Xung_100ms" THEN "Act_can_mau" := "Act_can_mau" + 1.12; END_IF;
   IF #_w1 THEN "TL_mau" := "Act_can_mau"; END_IF;
   IF "AlwaysTRUE" AND "Q_V2_Mau" AND "TG_Xung_100ms" THEN "Act_can_mau" := "Act_can_mau" - 1.3; END_IF;
END_REGION

REGION Network 5
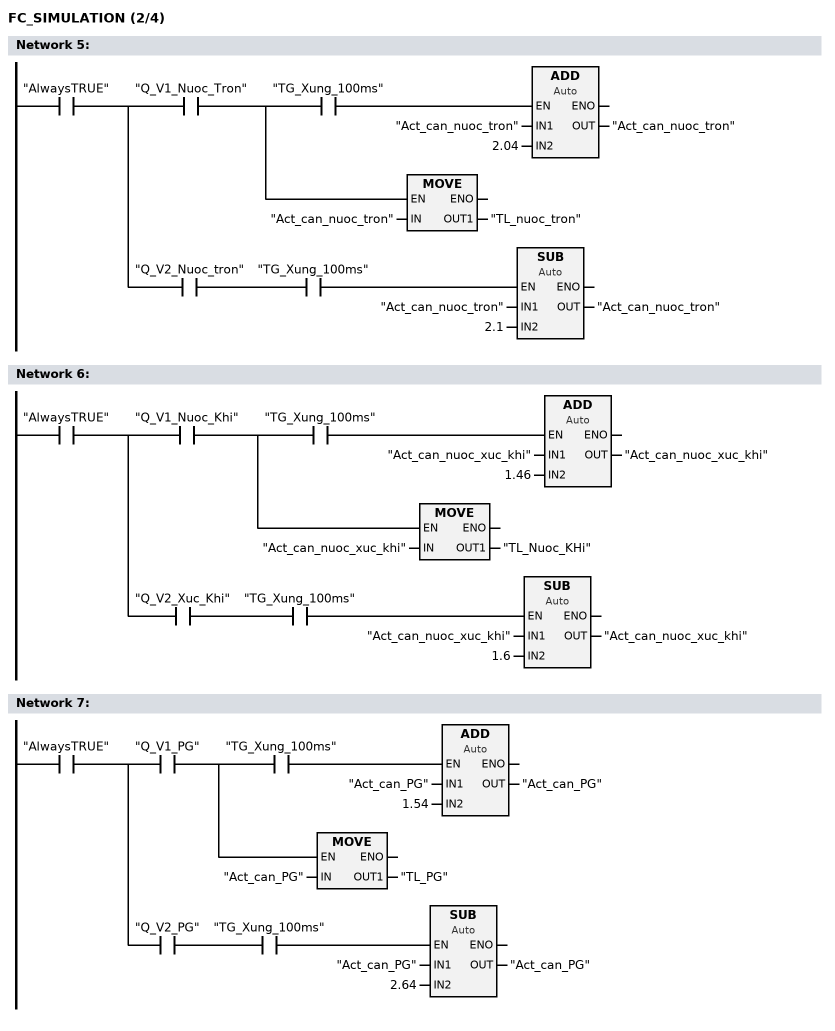
   RUNG wire#powerrail
      Contact( "AlwaysTRUE" )
      wire#w1
      Contact( "Q_V1_Nuoc_Tron" )
      wire#w2
      Contact( "TG_Xung_100ms" )
      Add(in1 := "Act_can_nuoc_tron", in2 := 2.04, out => "Act_can_nuoc_tron")
   END_RUNG
   RUNG wire#w2
      Move(in := "Act_can_nuoc_tron", out1 => "TL_nuoc_tron")
   END_RUNG
   RUNG wire#w1
      Contact( "Q_V2_Nuoc_tron" )
      Contact( "TG_Xung_100ms" )
      Sub(in1 := "Act_can_nuoc_tron", in2 := 2.1, out => "Act_can_nuoc_tron")
   END_RUNG
   // the same network as SCL:
   #_w1 := "AlwaysTRUE" AND "Q_V1_Nuoc_Tron";
   IF #_w1 AND "TG_Xung_100ms" THEN "Act_can_nuoc_tron" := "Act_can_nuoc_tron" + 2.04; END_IF;
   IF #_w1 THEN "TL_nuoc_tron" := "Act_can_nuoc_tron"; END_IF;
   IF "AlwaysTRUE" AND "Q_V2_Nuoc_tron" AND "TG_Xung_100ms" THEN
       "Act_can_nuoc_tron" := "Act_can_nuoc_tron" - 2.1;
   END_IF;
END_REGION

REGION Network 6
   RUNG wire#powerrail
      Contact( "AlwaysTRUE" )
      wire#w1
      Contact( "Q_V1_Nuoc_Khi" )
      wire#w2
      Contact( "TG_Xung_100ms" )
      Add(in1 := "Act_can_nuoc_xuc_khi", in2 := 1.46, out => "Act_can_nuoc_xuc_khi")
   END_RUNG
   RUNG wire#w2
      Move(in := "Act_can_nuoc_xuc_khi", out1 => "TL_Nuoc_KHi")
   END_RUNG
   RUNG wire#w1
      Contact( "Q_V2_Xuc_Khi" )
      Contact( "TG_Xung_100ms" )
      Sub(in1 := "Act_can_nuoc_xuc_khi", in2 := 1.6, out => "Act_can_nuoc_xuc_khi")
   END_RUNG
   // the same network as SCL:
   #_w1 := "AlwaysTRUE" AND "Q_V1_Nuoc_Khi";
   IF #_w1 AND "TG_Xung_100ms" THEN "Act_can_nuoc_xuc_khi" := "Act_can_nuoc_xuc_khi" + 1.46; END_IF;
   IF #_w1 THEN "TL_Nuoc_KHi" := "Act_can_nuoc_xuc_khi"; END_IF;
   IF "AlwaysTRUE" AND "Q_V2_Xuc_Khi" AND "TG_Xung_100ms" THEN
       "Act_can_nuoc_xuc_khi" := "Act_can_nuoc_xuc_khi" - 1.6;
   END_IF;
END_REGION

REGION Network 7
   RUNG wire#powerrail
      Contact( "AlwaysTRUE" )
      wire#w1
      Contact( "Q_V1_PG" )
      wire#w2
      Contact( "TG_Xung_100ms" )
      Add(in1 := "Act_can_PG", in2 := 1.54, out => "Act_can_PG")
   END_RUNG
   RUNG wire#w2
      Move(in := "Act_can_PG", out1 => "TL_PG")
   END_RUNG
   RUNG wire#w1
      Contact( "Q_V2_PG" )
      Contact( "TG_Xung_100ms" )
      Sub(in1 := "Act_can_PG", in2 := 2.64, out => "Act_can_PG")
   END_RUNG
   // the same network as SCL:
   #_w1 := "AlwaysTRUE" AND "Q_V1_PG";
   IF #_w1 AND "TG_Xung_100ms" THEN "Act_can_PG" := "Act_can_PG" + 1.54; END_IF;
   IF #_w1 THEN "TL_PG" := "Act_can_PG"; END_IF;
   IF "AlwaysTRUE" AND "Q_V2_PG" AND "TG_Xung_100ms" THEN "Act_can_PG" := "Act_can_PG" - 2.64; END_IF;
END_REGION

REGION Network 8: Bon 1
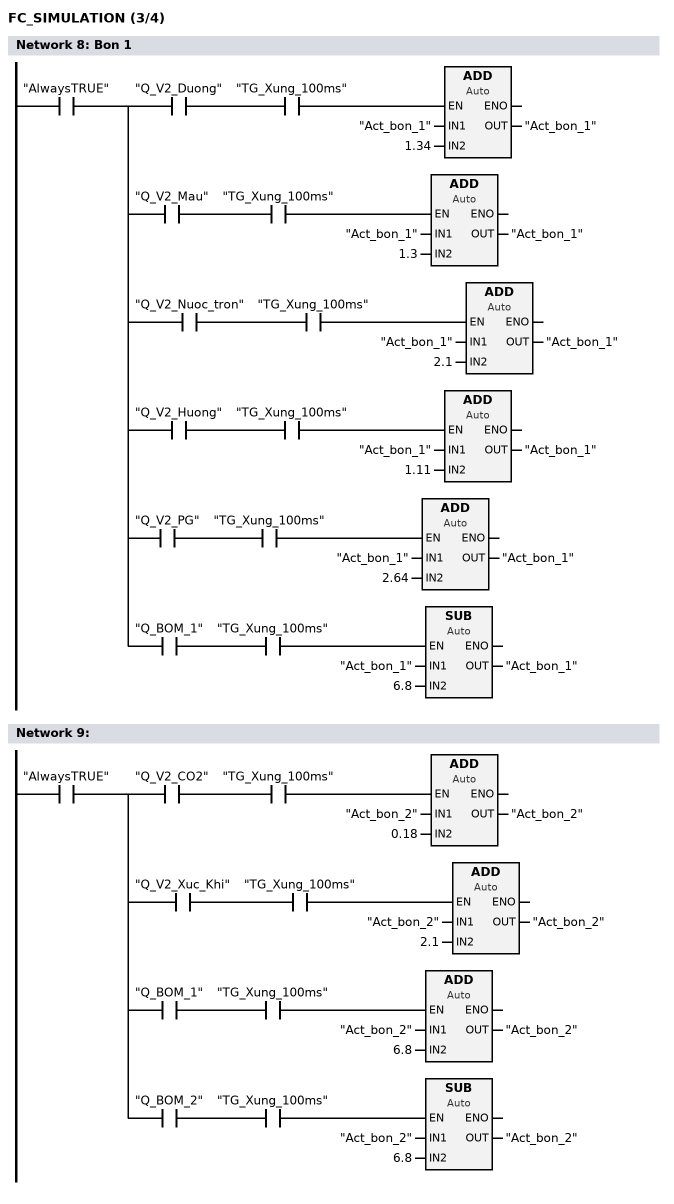
   RUNG wire#powerrail
      Contact( "AlwaysTRUE" )
      wire#w1
      Contact( "Q_V2_Duong" )
      Contact( "TG_Xung_100ms" )
      Add(in1 := "Act_bon_1", in2 := 1.34, out => "Act_bon_1")
   END_RUNG
   RUNG wire#w1
      Contact( "Q_V2_Mau" )
      Contact( "TG_Xung_100ms" )
      Add(in1 := "Act_bon_1", in2 := 1.3, out => "Act_bon_1")
   END_RUNG
   RUNG wire#w1
      Contact( "Q_V2_Nuoc_tron" )
      Contact( "TG_Xung_100ms" )
      Add(in1 := "Act_bon_1", in2 := 2.1, out => "Act_bon_1")
   END_RUNG
   RUNG wire#w1
      Contact( "Q_V2_Huong" )
      Contact( "TG_Xung_100ms" )
      Add(in1 := "Act_bon_1", in2 := 1.11, out => "Act_bon_1")
   END_RUNG
   RUNG wire#w1
      Contact( "Q_V2_PG" )
      Contact( "TG_Xung_100ms" )
      Add(in1 := "Act_bon_1", in2 := 2.64, out => "Act_bon_1")
   END_RUNG
   RUNG wire#w1
      Contact( "Q_BOM_1" )
      Contact( "TG_Xung_100ms" )
      Sub(in1 := "Act_bon_1", in2 := 6.8, out => "Act_bon_1")
   END_RUNG
   // the same network as SCL:
   IF "AlwaysTRUE" AND "Q_V2_Duong" AND "TG_Xung_100ms" THEN "Act_bon_1" := "Act_bon_1" + 1.34; END_IF;
   IF "AlwaysTRUE" AND "Q_V2_Mau" AND "TG_Xung_100ms" THEN "Act_bon_1" := "Act_bon_1" + 1.3; END_IF;
   IF "AlwaysTRUE" AND "Q_V2_Nuoc_tron" AND "TG_Xung_100ms" THEN "Act_bon_1" := "Act_bon_1" + 2.1; END_IF;
   IF "AlwaysTRUE" AND "Q_V2_Huong" AND "TG_Xung_100ms" THEN "Act_bon_1" := "Act_bon_1" + 1.11; END_IF;
   IF "AlwaysTRUE" AND "Q_V2_PG" AND "TG_Xung_100ms" THEN "Act_bon_1" := "Act_bon_1" + 2.64; END_IF;
   IF "AlwaysTRUE" AND "Q_BOM_1" AND "TG_Xung_100ms" THEN "Act_bon_1" := "Act_bon_1" - 6.8; END_IF;
END_REGION

REGION Network 9
   RUNG wire#powerrail
      Contact( "AlwaysTRUE" )
      wire#w1
      Contact( "Q_V2_CO2" )
      Contact( "TG_Xung_100ms" )
      Add(in1 := "Act_bon_2", in2 := 0.18, out => "Act_bon_2")
   END_RUNG
   RUNG wire#w1
      Contact( "Q_V2_Xuc_Khi" )
      Contact( "TG_Xung_100ms" )
      Add(in1 := "Act_bon_2", in2 := 2.1, out => "Act_bon_2")
   END_RUNG
   RUNG wire#w1
      Contact( "Q_BOM_1" )
      Contact( "TG_Xung_100ms" )
      Add(in1 := "Act_bon_2", in2 := 6.8, out => "Act_bon_2")
   END_RUNG
   RUNG wire#w1
      Contact( "Q_BOM_2" )
      Contact( "TG_Xung_100ms" )
      Sub(in1 := "Act_bon_2", in2 := 6.8, out => "Act_bon_2")
   END_RUNG
   // the same network as SCL:
   IF "AlwaysTRUE" AND "Q_V2_CO2" AND "TG_Xung_100ms" THEN "Act_bon_2" := "Act_bon_2" + 0.18; END_IF;
   IF "AlwaysTRUE" AND "Q_V2_Xuc_Khi" AND "TG_Xung_100ms" THEN "Act_bon_2" := "Act_bon_2" + 2.1; END_IF;
   IF "AlwaysTRUE" AND "Q_BOM_1" AND "TG_Xung_100ms" THEN "Act_bon_2" := "Act_bon_2" + 6.8; END_IF;
   IF "AlwaysTRUE" AND "Q_BOM_2" AND "TG_Xung_100ms" THEN "Act_bon_2" := "Act_bon_2" - 6.8; END_IF;
END_REGION

REGION Network 10
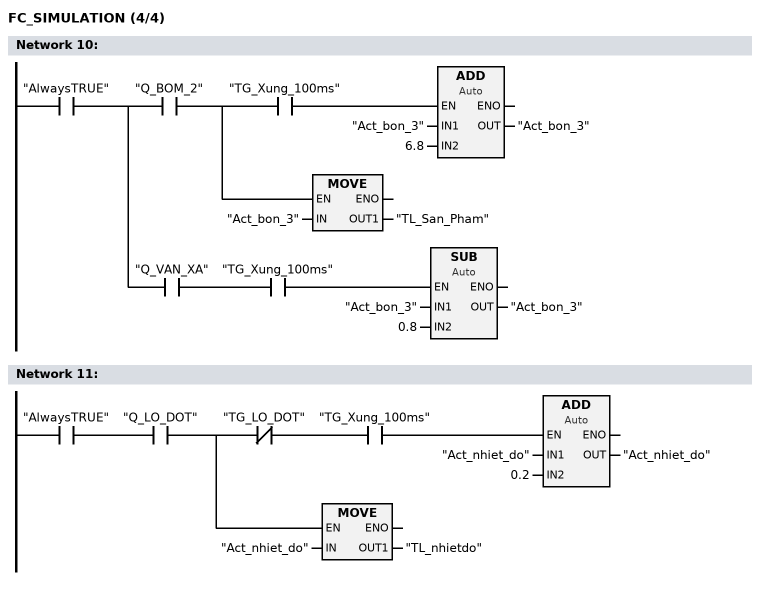
   RUNG wire#powerrail
      Contact( "AlwaysTRUE" )
      wire#w1
      Contact( "Q_BOM_2" )
      wire#w2
      Contact( "TG_Xung_100ms" )
      Add(in1 := "Act_bon_3", in2 := 6.8, out => "Act_bon_3")
   END_RUNG
   RUNG wire#w2
      Move(in := "Act_bon_3", out1 => "TL_San_Pham")
   END_RUNG
   RUNG wire#w1
      Contact( "Q_VAN_XA" )
      Contact( "TG_Xung_100ms" )
      Sub(in1 := "Act_bon_3", in2 := 0.8, out => "Act_bon_3")
   END_RUNG
   // the same network as SCL:
   #_w1 := "AlwaysTRUE" AND "Q_BOM_2";
   IF #_w1 AND "TG_Xung_100ms" THEN "Act_bon_3" := "Act_bon_3" + 6.8; END_IF;
   IF #_w1 THEN "TL_San_Pham" := "Act_bon_3"; END_IF;
   IF "AlwaysTRUE" AND "Q_VAN_XA" AND "TG_Xung_100ms" THEN "Act_bon_3" := "Act_bon_3" - 0.8; END_IF;
END_REGION

REGION Network 11
   RUNG wire#powerrail
      Contact( "AlwaysTRUE" )
      Contact( "Q_LO_DOT" )
      wire#w1
      I_Contact( "TG_LO_DOT" )
      Contact( "TG_Xung_100ms" )
      Add(in1 := "Act_nhiet_do", in2 := 0.2, out => "Act_nhiet_do")
   END_RUNG
   RUNG wire#w1
      Move(in := "Act_nhiet_do", out1 => "TL_nhietdo")
   END_RUNG
   // the same network as SCL:
   #_w1 := "AlwaysTRUE" AND "Q_LO_DOT";
   IF #_w1 AND NOT "TG_LO_DOT" AND "TG_Xung_100ms" THEN "Act_nhiet_do" := "Act_nhiet_do" + 0.2; END_IF;
   IF #_w1 THEN "TL_nhietdo" := "Act_nhiet_do"; END_IF;
END_REGION
END_FUNCTION

ORGANIZATION_BLOCK "Main"   // OB1, LAD, ProgramCycle
TITLE = "Main Program Sweep (Cycle)"
{ S7_Optimized_Access := 'TRUE' }
VERSION : 0.1
   VAR_INPUT
      Initial_Call : Bool;   // Initial call of this OB
      Remanence : Bool;   // =True, if remanent data are available
   END_VAR
   VAR_TEMP   // added for the SCL form of the ladder/FBD networks
      _w1 : Bool;
   END_VAR
BEGIN

REGION Network 1: Chọn Chế Độ
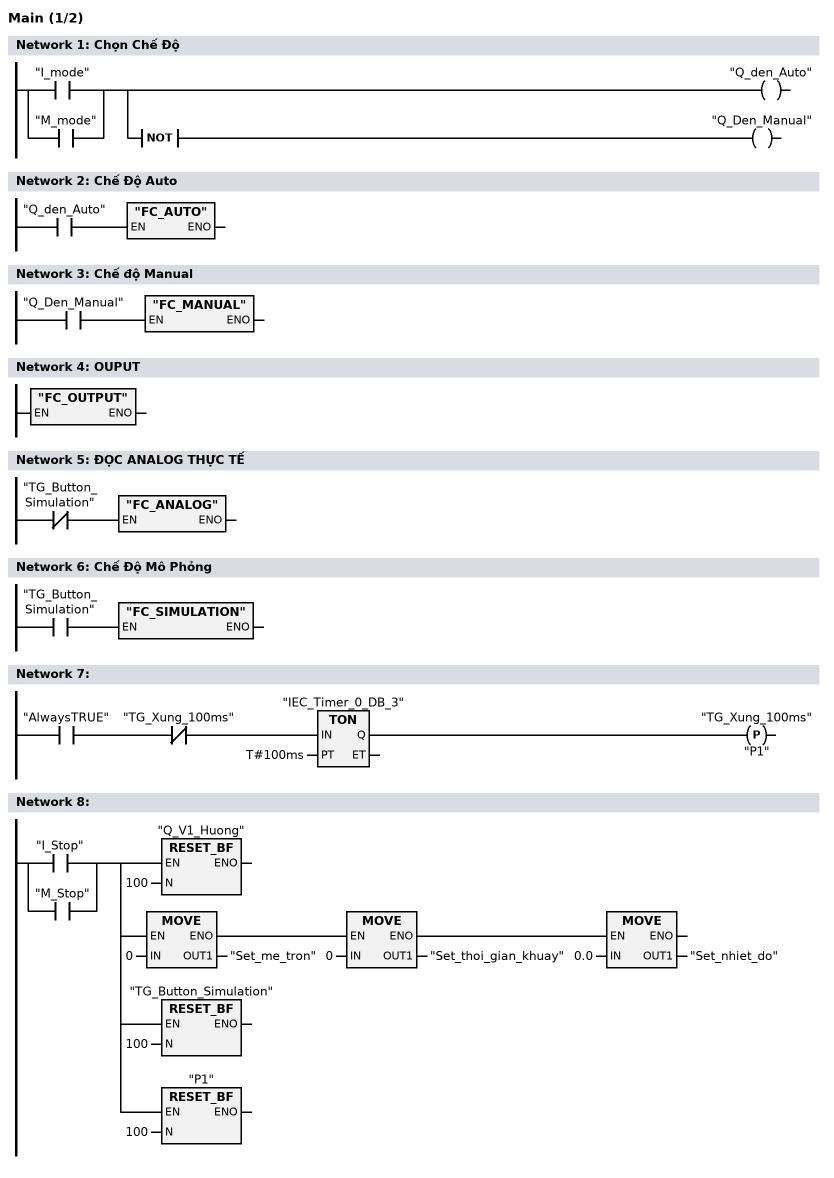
   RUNG wire#powerrail
      Contact( "I_mode" )
      wire#w1
      Coil( "Q_den_Auto" )
   END_RUNG
   RUNG wire#powerrail
      Contact( "M_mode" )
   END_RUNG wire#w1
   RUNG wire#w1
      Not()
      Coil( "Q_Den_Manual" )
   END_RUNG
   // the same network as SCL:
   "Q_den_Auto" := "I_mode" OR "M_mode";
   "Q_Den_Manual" := NOT "Q_den_Auto";
END_REGION

REGION Network 2: Chế Độ Auto
   RUNG wire#powerrail
      Contact( "Q_den_Auto" )
      "FC_AUTO"()
   END_RUNG
   // the same network as SCL:
   IF "Q_den_Auto" THEN "FC_AUTO"(); END_IF;
END_REGION

REGION Network 3: Chế độ Manual
   RUNG wire#powerrail
      Contact( "Q_Den_Manual" )
      "FC_MANUAL"()
   END_RUNG
   // the same network as SCL:
   IF "Q_Den_Manual" THEN "FC_MANUAL"(); END_IF;
END_REGION

REGION Network 4: OUPUT
   RUNG wire#powerrail
      "FC_OUTPUT"()
   END_RUNG
   // the same network as SCL:
   "FC_OUTPUT"();
END_REGION

REGION Network 5: ĐỌC ANALOG THỰC TẾ
   RUNG wire#powerrail
      I_Contact( "TG_Button_Simulation" )
      "FC_ANALOG"()
   END_RUNG
   // the same network as SCL:
   IF NOT "TG_Button_Simulation" THEN "FC_ANALOG"(); END_IF;
END_REGION

REGION Network 6: Chế Độ Mô Phỏng
   RUNG wire#powerrail
      Contact( "TG_Button_Simulation" )
      "FC_SIMULATION"()
   END_RUNG
   // the same network as SCL:
   IF "TG_Button_Simulation" THEN "FC_SIMULATION"(); END_IF;
END_REGION

REGION Network 7
   "IEC_Timer_0_DB_3".TON(IN := "AlwaysTRUE" AND NOT "TG_Xung_100ms", PT := T#100ms);
   "TG_Xung_100ms" := "IEC_Timer_0_DB_3".Q AND NOT "P1";   // rising edge
   "P1" := "IEC_Timer_0_DB_3".Q;
END_REGION

REGION Network 8
   // no SCL statement known for RBitfield: written as a call
   #_w1 := "I_Stop" OR "M_Stop";
   IF #_w1 THEN
       RESET_BF(operand := "Q_V1_Huong", n := 100);
       "Set_me_tron" := 0;
       "Set_thoi_gian_khuay" := 0;
       "Set_nhiet_do" := 0.0;
       RESET_BF(operand := "TG_Button_Simulation", n := 100);
       RESET_BF(operand := "P1", n := 100);
   END_IF;
END_REGION

REGION Network 9
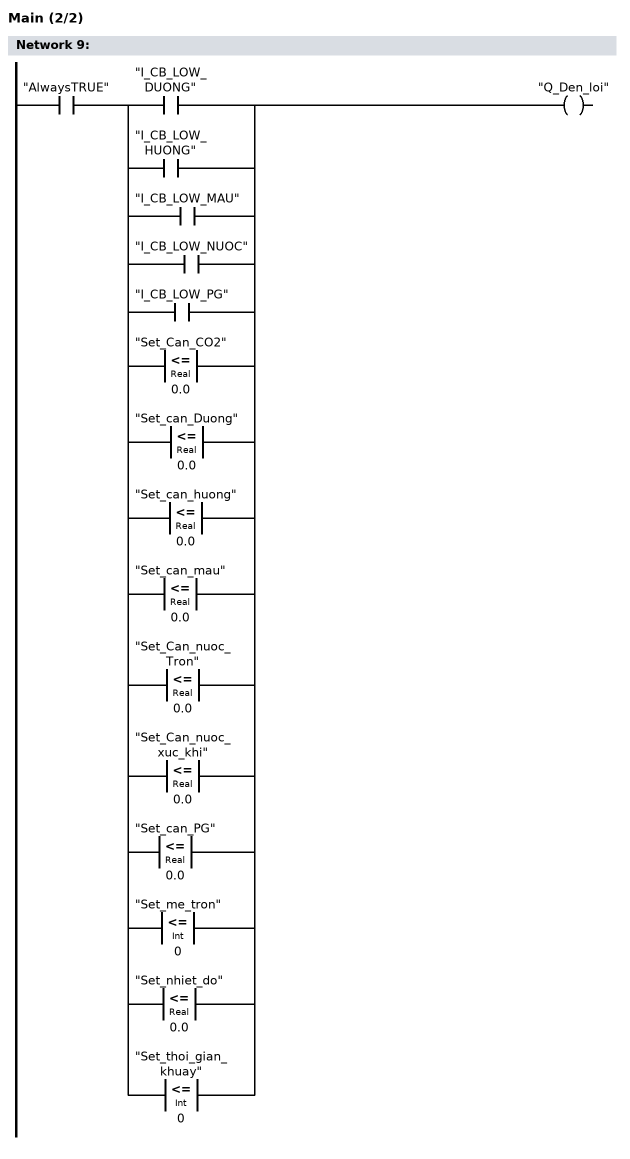
   RUNG wire#powerrail
      Contact( "AlwaysTRUE" )
      wire#w1
      Contact( "I_CB_LOW_DUONG" )
      wire#w2
      Coil( "Q_Den_loi" )
   END_RUNG
   RUNG wire#w1
      Contact( "I_CB_LOW_HUONG" )
   END_RUNG wire#w2
   RUNG wire#w1
      Contact( "I_CB_LOW_MAU" )
   END_RUNG wire#w2
   RUNG wire#w1
      Contact( "I_CB_LOW_NUOC" )
   END_RUNG wire#w2
   RUNG wire#w1
      Contact( "I_CB_LOW_PG" )
   END_RUNG wire#w2
   RUNG wire#w1
      { S7_Templates := "SrcType := Real" } LE_Contact(in1 := "Set_Can_CO2", in2 := 0.0)
   END_RUNG wire#w2
   RUNG wire#w1
      { S7_Templates := "SrcType := Real" } LE_Contact(in1 := "Set_can_Duong", in2 := 0.0)
   END_RUNG wire#w2
   RUNG wire#w1
      { S7_Templates := "SrcType := Real" } LE_Contact(in1 := "Set_can_huong", in2 := 0.0)
   END_RUNG wire#w2
   RUNG wire#w1
      { S7_Templates := "SrcType := Real" } LE_Contact(in1 := "Set_can_mau", in2 := 0.0)
   END_RUNG wire#w2
   RUNG wire#w1
      { S7_Templates := "SrcType := Real" } LE_Contact(in1 := "Set_Can_nuoc_Tron", in2 := 0.0)
   END_RUNG wire#w2
   RUNG wire#w1
      { S7_Templates := "SrcType := Real" } LE_Contact(in1 := "Set_Can_nuoc_xuc_khi", in2 := 0.0)
   END_RUNG wire#w2
   RUNG wire#w1
      { S7_Templates := "SrcType := Real" } LE_Contact(in1 := "Set_can_PG", in2 := 0.0)
   END_RUNG wire#w2
   RUNG wire#w1
      { S7_Templates := "SrcType := Int" } LE_Contact(in1 := "Set_me_tron", in2 := 0)
   END_RUNG wire#w2
   RUNG wire#w1
      { S7_Templates := "SrcType := Real" } LE_Contact(in1 := "Set_nhiet_do", in2 := 0.0)
   END_RUNG wire#w2
   RUNG wire#w1
      { S7_Templates := "SrcType := Int" } LE_Contact(in1 := "Set_thoi_gian_khuay", in2 := 0)
   END_RUNG wire#w2
   // the same network as SCL:
   "Q_Den_loi" := "AlwaysTRUE" AND ("I_CB_LOW_DUONG" OR "I_CB_LOW_HUONG" OR "I_CB_LOW_MAU" OR "I_CB_LOW_NUOC" OR "I_CB_LOW_PG" OR ("Set_Can_CO2" <= 0.0) OR ("Set_can_Duong" <= 0.0) OR ("Set_can_huong" <= 0.0) OR ("Set_can_mau" <= 0.0) OR ("Set_Can_nuoc_Tron" <= 0.0) OR ("Set_Can_nuoc_xuc_khi" <= 0.0) OR ("Set_can_PG" <= 0.0) OR ("Set_me_tron" <= 0) OR ("Set_nhiet_do" <= 0.0) OR ("Set_thoi_gian_khuay" <= 0));
END_REGION
END_ORGANIZATION_BLOCK

(* ===== HMI "HMI_RT_1" =====
system functions are stored by id; their names below are inferred from use
connection "HMI_Connection_1": ETHERNET, S7_1200_OMS
connection "HMI_Connection_2": ETHERNET, S7_1200_OMS

HMI tags "Default tag table"
   "M_CB_LOW_HUONG" : Bool = PLC M_CB_LOW_HUONG AT %M13.0, 1 s
   "M_CB_LOW_MAU" : Bool = PLC M_CB_LOW_MAU AT %M13.1, 1 s
   "M_CB_LOW_PG" : Bool = PLC M_CB_LOW_PG AT %M13.2, 1 s
   "M_CB_LOW_NUOC" : Bool = PLC M_CB_LOW_NUOC AT %M13.4, 1 s
   "M_CB_LOW_CO2" : Real = PLC M_CB_LOW_CO2 AT %MD500, 1 s
   "M_CB_LOW_BON_2" : Real = PLC M_CB_LOW_BON_2 AT %MD504, 1 s
   "M_CB_CHAI" : Bool = PLC M_CB_CHAI AT %M13.7, 1 s
   "Q_V1_Huong" : Bool = PLC Q_V1_Huong AT %Q0.3, 1 s
   "Q_V2_Huong" : Bool = PLC Q_V2_Huong AT %Q0.4, 1 s
   "Q_V1_Mau" : Bool = PLC Q_V1_Mau AT %Q0.5, 1 s
   "Q_V2_Mau" : Bool = PLC Q_V2_Mau AT %Q0.6, 1 s
   "Q_V1_PG" : Bool = PLC Q_V1_PG AT %Q0.7, 1 s
   "Q_V2_PG" : Bool = PLC Q_V2_PG AT %Q1.0, 1 s
   "Q_V1_Duong" : Bool = PLC Q_V1_Duong AT %Q1.3, 1 s
   "M_CB_LOW_DUONG" : Bool = PLC M_CB_LOW_DUONG AT %M13.3, 1 s
   "Q_V2_Duong" : Bool = PLC Q_V2_Duong AT %Q1.4, 1 s
   "Q_V1_Nuoc_Tron" : Bool = PLC Q_V1_Nuoc_Tron AT %Q1.1, 1 s
   "Q_V2_Nuoc_tron" : Bool = PLC Q_V2_Nuoc_tron AT %Q1.2, 1 s
   "Q_V1_Nuoc_Khi" : Bool = PLC Q_V1_Nuoc_Khi AT %Q1.5, 1 s
   "Q_V2_Xuc_Khi" : Bool = PLC Q_V2_Xuc_Khi AT %Q1.6, 1 s
   "Q_V1_CO2" : Bool = PLC Q_V1_CO2 AT %Q1.7, 1 s
   "Q_V2_CO2" : Bool = PLC Q_V2_CO2 AT %Q2.0, 1 s
   "Q_BOM_1" : Bool = PLC Q_BOM_1 AT %Q2.3, 1 s
   "Q_BOM_2" : Bool = PLC Q_BOM_2 AT %Q2.4, 1 s
   "Q_BOM_TRON" : Bool = PLC Q_BOM_TRON AT %Q2.1, 1 s
   "Q_VAN_XA" : Bool = PLC Q_VAN_XA AT %Q2.5, 1 s
   "Q_BT" : Bool = PLC Q_BT AT %Q2.7, 1 s
   "M_SW_V1_Huong" : Bool = PLC M_SW_V1_Huong AT %M10.3, 1 s
   "M_SW_V1_mau" : Bool = PLC M_SW_V1_mau AT %M10.5, 1 s
   "M_SW_V1_PG" : Bool = PLC M_SW_V1_PG AT %M10.7, 1 s
   "M_SW_V1_Nuoc_Tron" : Bool = PLC M_SW_V1_Nuoc_Tron AT %M11.3, 1 s
   "M_SW_V1_Nuoc_Xuc_Khi" : Bool = PLC M_SW_V1_Nuoc_Xuc_Khi AT %M11.5, 1 s
   "M_SW_V1_CO2" : Bool = PLC M_SW_V1_CO2 AT %M11.7, 1 s
   "M_SW_V1_Duong" : Bool = PLC M_SW_V1_Duong AT %M11.1, 1 s
   "M_SW_V2_Huong" : Bool = PLC M_SW_V2_Huong AT %M10.4, 1 s
   "M_SW_V2_mau" : Bool = PLC M_SW_V2_mau AT %M10.6, 1 s
   "M_SW_V2_PG" : Bool = PLC M_SW_V2_PG AT %M11.0, 1 s
   "M_SW_V2_Duong" : Bool = PLC M_SW_V2_Duong AT %M11.2, 1 s
   "M_SW_V2_Nuoc_Tron" : Bool = PLC M_SW_V2_Nuoc_Tron AT %M11.4, 1 s
   "M_SW_V2_Nuoc_Xuc_Khi" : Bool = PLC M_SW_V2_Nuoc_Xuc_Khi AT %M11.6, 1 s
   "M_SW_V2_CO2" : Bool = PLC M_SW_V2_CO2 AT %M12.0, 1 s
   "M_SW_BOM_TRON" : Bool = PLC M_SW_BOM_TRON AT %M12.1, 1 s
   "M_SW_LAM_LANH" : Bool = PLC M_SW_LAM_LANH AT %M12.2, 1 s
   "M_SW_LO_DOT" : Bool = PLC M_SW_LO_DOT AT %M12.5, 1 s
   "M_SW_BOM_1" : Bool = PLC M_SW_BOM_1 AT %M12.3, 1 s
   "M_SW_BOM_2" : Bool = PLC M_SW_BOM_2 AT %M12.4, 1 s
   "M_SW_VAN_XA" : Bool = PLC M_SW_VAN_XA AT %M12.6, 1 s
   "Q_LO_DOT" : Bool = PLC Q_LO_DOT AT %Q2.6, 1 s
   "M_mode" : Bool = PLC M_mode AT %M10.0, 1 s
   "M_start" : Bool = PLC M_start AT %M10.1, 1 s
   "M_Stop" : Bool = PLC M_Stop AT %M10.2, 1 s
   "TG_Button_Simulation" : Bool = PLC TG_Button_Simulation AT %M40.0, 1 s
   "TG_DK_RUN" : Bool = PLC TG_DK_RUN AT %M41.0, 1 s
   "Q_Den_loi" : Bool = PLC Q_Den_loi AT %Q0.2, 1 s
   "Q_Den_Manual" : Bool = PLC Q_Den_Manual AT %Q0.1, 1 s
   "Q_den_Auto" : Bool = PLC Q_den_Auto AT %Q0.0, 1 s
   "Act_time_Khuay" : Int = PLC Act_time_Khuay AT %MW400, 1 s
   "Act_nhiet_do" : Real = PLC Act_nhiet_do AT %MD402, 1 s
   "Act_CO2" : Real = PLC Act_Can_CO2 AT %MD432, 1 s
   "Act_can_huong" : Real = PLC Act_can_huong AT %MD408, 1 s
   "Act_can_PG" : Real = PLC Act_can_PG AT %MD420, 1 s
   "Act_can_mau" : Real = PLC Act_can_mau AT %MD412, 1 s
   "Act_nuoc_tron" : Real = PLC Act_can_nuoc_tron AT %MD424, 1 s
   "Act_nuoc_xuc_khi" : Real = PLC Act_can_nuoc_xuc_khi AT %MD428, 1 s
   "Act_me" : Int = PLC Act_me AT %MW406, 1 s
   "Act_San_luong" : Int = PLC Act_So_chai AT %MW436, 1 s
   "Set_can_Duong" : Real = PLC Set_can_Duong AT %MD212, 1 s
   "Set_Can_CO2" : Real = PLC Set_Can_CO2 AT %MD224, 1 s
   "Set_can_huong" : Real = PLC Set_can_huong AT %MD200, 1 s
   "Set_can_mau" : Real = PLC Set_can_mau AT %MD204, 1 s
   "Set_Can_nuoc_Tron" : Real = PLC Set_Can_nuoc_Tron AT %MD216, 1 s
   "Set_Can_nuoc_xuc_khi" : Real = PLC Set_Can_nuoc_xuc_khi AT %MD220, 1 s
   "Set_can_PG" : Real = PLC Set_can_PG AT %MD208, 1 s
   "M_SW_BANG_TAI" : Bool = PLC M_SW_BANG_TAI AT %M12.7, 1 s
   "Act_can_duong" : Real = PLC Act_can_duong AT %MD416, 1 s
   "Q_LAM_LANH" : Bool = PLC Q_LAM_LANH AT %Q2.2, 1 s
   "Act_bon_1" : Real = PLC Act_bon_1 AT %MD440, 1 s
   "Act_bon_2" : Real = PLC Act_bon_2 AT %MD444, 1 s
   "Act_bon_3" : Real = PLC Act_bon_3 AT %MD448, 1 s
   "TL_San_Pham" : Real = PLC TL_San_Pham AT %MD628, 1 s
   "TL_CO2" : Real = PLC TL_CO2 AT %MD620, 1 s
   "TL_Nuoc_KHi" : Real = PLC TL_Nuoc_KHi AT %MD624, 1 s
   "TL_nuoc_tron" : Real = PLC TL_nuoc_tron AT %MD616, 1 s
   "TL_mau" : Real = PLC TL_mau AT %MD604, 1 s
   "TL_PG" : Real = PLC TL_PG AT %MD612, 1 s
   "TL_Huong" : Real = PLC TL_Huong AT %MD600, 1 s
   "TL_nhietdo" : Real = PLC TL_nhietdo AT %MD636, 1 s
   "TL_thoiGian_khuay" : DInt = PLC TL_thoiGian_khuay AT %MD632, 1 s
   "TL_Duong" : Real = PLC TL_Duong AT %MD608, 1 s
   "TG_VT_SP" : DInt = PLC TG_VT_SP AT %MD508, 1 s
   "Tag_Dang_nhap" : WString[254] AT %DB1.DBX0.0
   "Set_thoi_gian_khuay" : Int = PLC Set_thoi_gian_khuay AT %MW228, 1 s
   "Set_me_tron" : Int = PLC Set_me_tron AT %MW304, 1 s
   "Set_nhiet_do" : Real = PLC Set_nhiet_do AT %MD300, 1 s
   "User_Input" : WString[50], internal
   "Pass_Input" : WString[50], internal
   "Login_Status" : WString[50], internal

screen "Screen_1" 1600x1200
   SymbolLibrary "Symbol library_95" at 1030,723 size 9x40
      Appearance <- "Q_VAN_XA"
   SymbolLibrary "Symbol library_87" at 695,545 size 16x19
      Appearance <- "Q_V2_CO2"
   SymbolLibrary "Symbol library_75" at 784,480 size 9x42
      Appearance <- "Q_V2_Xuc_Khi"
   SymbolLibrary "Symbol library_61" at 495,485 size 9x25
      Appearance <- "Q_V2_Duong"
   SymbolLibrary "Symbol library_58" at 318,490 size 58x9
      Appearance <- "Q_V2_PG"
   SymbolLibrary "Symbol library_57" at 368,479 size 16x19
      Appearance <- "Q_V2_PG"
   SymbolLibrary "Symbol library_55" at 214,478 size 9x85
      Appearance <- "Q_V2_Mau"
   SymbolLibrary "Symbol library_54" at 186,503 size 9x64
      Appearance <- "Q_V2_Huong"
   SymbolLibrary "Symbol library_50" at 784,387 size 9x57
      Appearance <- "Q_V2_Xuc_Khi"
   SymbolLibrary "Symbol library_49" at 788,257 size 9x57
      Appearance <- "Q_V1_Nuoc_Khi"
   SymbolLibrary "Symbol library_44" at 661,385 size 9x48
      Appearance <- "Q_V2_Nuoc_tron"
   SymbolLibrary "Symbol library_43" at 662,126 size 16x19
      Appearance <- "Q_V1_Nuoc_Tron"
   SymbolLibrary "Symbol library_42" at 663,262 size 9x55
      Appearance <- "Q_V1_Nuoc_Tron"
   SymbolLibrary "Symbol library_41" at 662,144 size 9x75
      Appearance <- "Q_V1_Nuoc_Tron"
   SymbolLibrary "Symbol library_40" at 495,389 size 9x56
      Appearance <- "Q_V2_Duong"
   SymbolLibrary "Symbol library_39" at 496,199 size 9x113
      Appearance <- "Q_V1_Duong"
   SymbolLibrary "Symbol library_36" at 373,385 size 9x56
      Appearance <- "Q_V2_PG"
   SymbolLibrary "Symbol library_35" at 373,257 size 9x56
      Appearance <- "Q_V1_PG"
   SymbolLibrary "Symbol library_34" at 372,178 size 9x45
      Appearance <- "Q_V1_PG"
   SymbolLibrary "Symbol library_33" at 221,263 size 9x51
      Appearance <- "Q_V1_Mau"
   SymbolLibrary "Symbol library_31" at 222,181 size 9x45
      Appearance <- "Q_V1_Mau"
   SymbolLibrary "Symbol library_30" at 215,388 size 9x52
      Appearance <- "Q_V2_Mau"
   SymbolLibrary "Symbol library_32" at 78,180 size 9x41
      Appearance <- "Q_V1_Huong"
   GraphicView "Graphic view_1" at 9,3 size 57x56; Picture "UTC2"
   TextField "Text field_1" at 85,14 size 547x24; Text 'HỆ THỐNG SCADA CHO DÂY CHUYỀN SẢN XUẤT NƯỚC NGỌT'
   SymbolLibrary "Symbol library_56" at 41,97 size 86x87
   SymbolLibrary "Symbol library_24" at 34,218 size 59x46
      Appearance <- "Q_V1_Huong"
   SymbolLibrary "Symbol library_1" at 183,97 size 86x87
   SymbolLibrary "Symbol library_2" at 335,99 size 86x87
   SymbolLibrary "Symbol library_4" at 177,222 size 59x46
      Appearance <- "Q_V1_Mau"
   SymbolLibrary "Symbol library_5" at 328,215 size 59x46
      Appearance <- "Q_V1_PG"
   SymbolLibrary "Symbol library_8" at 52,314 size 60x80
   SymbolLibrary "Symbol library_6" at 189,311 size 60x80
   SymbolLibrary "Symbol library_7" at 347,307 size 60x80
   SymbolLibrary "Symbol library_9" at 471,311 size 60x80
   SymbolLibrary "Symbol library_25" at 32,431 size 60x55
      Appearance <- "Q_V2_Huong"
   SymbolLibrary "Symbol library_10" at 169,424 size 60x55
      Appearance <- "Q_V2_Mau"
   SymbolLibrary "Symbol library_11" at 328,427 size 60x55
      Appearance <- "Q_V2_PG"
   SymbolLibrary "Symbol library_12" at 518,183 size 80x71
   SymbolLibrary "Symbol library_3" at 518,81 size 84x134
   SymbolLibrary "Symbol library_18" at 569,165 size 68x50
      Appearance <- "Q_V1_Duong"
   SymbolLibrary "Symbol library_13" at 449,431 size 60x55
      Appearance <- "Q_V2_Duong"
   IOField "I/O field_3" at 106,288 size 78x32; FormatPattern 999999999.999
      ProcessValue <- "Act_can_huong"
   IOField "I/O field_1" at 249,288 size 78x32; FormatPattern 999999999.999
      ProcessValue <- "Act_can_mau"
   IOField "I/O field_2" at 402,278 size 78x32; FormatPattern 999999999.999
      ProcessValue <- "Act_can_PG"
   IOField "I/O field_4" at 509,277 size 78x32; FormatPattern 999999999.999
      ProcessValue <- "Act_can_duong"
   SymbolLibrary "Symbol library_14" at 179,555 size 191x175
   SymbolLibrary "Symbol library_15" at 184,719 size 183x108
   SymbolLibrary "Symbol library_64" at 184,720 size 183x108
      Visibility <- "Q_LO_DOT"
   SymbolLibrary "Symbol library_21" at 223,473 size 104x222
      Appearance <- "Q_BOM_TRON"
   SymbolLibrary "Symbol library_16" at 675,81 size 105x115
   SymbolLibrary "Symbol library_17" at 618,217 size 59x46
      Appearance <- "Q_V1_Nuoc_Tron"
   SymbolLibrary "Symbol library_19" at 636,314 size 60x80
   SymbolLibrary "Symbol library_20" at 877,75 size 106x116
   SymbolLibrary "Symbol library_22" at 881,221 size 59x46
      Appearance <- "Q_V1_CO2"
   SymbolLibrary "Symbol library_23" at 898,324 size 60x80
   SymbolLibrary "Symbol library_26" at 614,421 size 60x55
      Appearance <- "Q_V2_Nuoc_tron"
   SymbolLibrary "Symbol library_27" at 738,428 size 60x55
      Appearance <- "Q_V2_Xuc_Khi"
   SymbolLibrary "Symbol library_28" at 79,263 size 9x52
      Appearance <- "Q_V1_Huong"
   SymbolLibrary "Symbol library_29" at 78,393 size 9x52
      Appearance <- "Q_V2_Huong"
   SymbolLibrary "Symbol library_37" at 507,182 size 76x9
      Appearance <- "Q_V1_Duong"
   SymbolLibrary "Symbol library_38" at 496,181 size 16x19
      Appearance <- "Q_V1_Duong"
   SymbolLibrary "Symbol library_45" at 743,214 size 59x46
      Appearance <- "Q_V1_Nuoc_Khi"
   SymbolLibrary "Symbol library_46" at 778,126 size 19x16
      Appearance <- "Q_V1_Nuoc_Khi"
   SymbolLibrary "Symbol library_47" at 788,141 size 9x75
      Appearance <- "Q_V1_Nuoc_Khi"
   SymbolLibrary "Symbol library_48" at 760,314 size 60x80
   SymbolLibrary "Symbol library_51" at 77,484 size 19x16
      Appearance <- "Q_V2_Huong"
   SymbolLibrary "Symbol library_52" at 88,492 size 90x9
      Appearance <- "Q_V2_Huong"
   SymbolLibrary "Symbol library_53" at 176,492 size 19x16
      Appearance <- "Q_V2_Huong"
   IOField "I/O field_5" at 688,275 size 78x32; FormatPattern 999999999.999
      ProcessValue <- "Act_nuoc_tron"
   IOField "I/O field_6" at 808,278 size 78x32; FormatPattern 999999999.999
      ProcessValue <- "Act_nuoc_xuc_khi"
   IOField "I/O field_7" at 961,283 size 78x32; FormatPattern 999999999.999
      ProcessValue <- "Act_CO2"
   SymbolLibrary "Symbol library_59" at 309,489 size 16x19
      Appearance <- "Q_V2_PG"
   SymbolLibrary "Symbol library_60" at 309,502 size 9x56
      Appearance <- "Q_V2_PG"
   SymbolLibrary "Symbol library_62" at 487,498 size 16x19
      Appearance <- "Q_V2_Duong"
   SymbolLibrary "Symbol library_63" at 334,508 size 159x9
      Appearance <- "Q_V2_Duong"
   SymbolLibrary "Symbol library_65" at 327,507 size 16x19
      Appearance <- "Q_V2_Duong"
   SymbolLibrary "Symbol library_66" at 327,521 size 9x39
      Appearance <- "Q_V2_Duong"
   SymbolLibrary "Symbol library_67" at 660,476 size 9x42
      Appearance <- "Q_V2_Nuoc_tron"
   SymbolLibrary "Symbol library_68" at 653,512 size 16x19
      Appearance <- "Q_V2_Nuoc_tron"
   SymbolLibrary "Symbol library_69" at 347,522 size 308x9
      Appearance <- "Q_V2_Nuoc_tron"
   SymbolLibrary "Symbol library_70" at 339,521 size 16x19
      Appearance <- "Q_V2_Nuoc_tron"
   SymbolLibrary "Symbol library_71" at 339,529 size 9x32
      Appearance <- "Q_V2_Nuoc_tron"
   SymbolLibrary "Symbol library_72" at 366,662 size 56x33
      Appearance <- "Q_BOM_1"
   SymbolLibrary "Symbol library_73" at 421,673 size 142x9
      Appearance <- "Q_BOM_1"
   SymbolLibrary "Symbol library_74" at 559,555 size 191x175
   SymbolLibrary "Symbol library_76" at 775,517 size 18x19
      Appearance <- "Q_V2_Xuc_Khi"
   SymbolLibrary "Symbol library_77" at 685,527 size 105x9
      Appearance <- "Q_V2_Xuc_Khi"
   SymbolLibrary "Symbol library_78" at 674,527 size 16x19
      Appearance <- "Q_V2_Xuc_Khi"
   SymbolLibrary "Symbol library_79" at 674,538 size 9x20
      Appearance <- "Q_V2_Xuc_Khi"
   SymbolLibrary "Symbol library_80" at 925,190 size 9x32
      Appearance <- "Q_V1_CO2"
   SymbolLibrary "Symbol library_81" at 925,266 size 9x59
      Appearance <- "Q_V1_CO2"
   SymbolLibrary "Symbol library_82" at 924,403 size 9x41
      Appearance <- "Q_V2_CO2"
   SymbolLibrary "Symbol library_83" at 879,430 size 60x55
      Appearance <- "Q_V2_CO2"
   SymbolLibrary "Symbol library_84" at 925,484 size 9x54
      Appearance <- "Q_V2_CO2"
   SymbolLibrary "Symbol library_85" at 916,536 size 18x19
      Appearance <- "Q_V2_CO2"
   SymbolLibrary "Symbol library_86" at 704,545 size 220x9
      Appearance <- "Q_V2_CO2"
   SymbolLibrary "Symbol library_88" at 748,662 size 56x33
      Appearance <- "Q_BOM_2"
   SymbolLibrary "Symbol library_89" at 939,551 size 191x175
   SymbolLibrary "Symbol library_90" at 804,672 size 138x9
      Appearance <- "Q_BOM_2"
   SymbolLibrary "Symbol library_91" at 481,622 size 50x40
   SymbolLibrary "Symbol library_92" at 527,646 size 37x6
      Appearance <- "Q_LAM_LANH"
   SymbolLibrary "Symbol library_93" at 527,654 size 37x6
      Appearance <- "Q_LAM_LANH"
   Bar "Bar_1" at 183,566 size 27x139; MinimumValue 0; MaximumValue 1000
      ProcessValue <- "Act_bon_1"
   Bar "Bar_2" at 715,565 size 32x139; MinimumValue 0; MaximumValue 1000
      ProcessValue <- "Act_bon_2"
   Bar "Bar_3" at 1100,559 size 27x139; MinimumValue 0; MaximumValue 1000
      ProcessValue <- "Act_bon_3"
   SymbolLibrary "Symbol library_94" at 984,749 size 60x55
      Appearance <- "Q_VAN_XA"
   SymbolLibrary "Symbol library_97" at 1022,802 size 17x19
      Appearance <- "Q_VAN_XA"
   SymbolLibrary "Symbol library_98" at 545,875 size 509x80
      Appearance <- "Q_BT"
   SymbolLibrary "Symbol library_99" at 866,812 size 159x9
      Appearance <- "Q_VAN_XA"
   SymbolLibrary "Symbol library_100" at 857,812 size 16x17
      Appearance <- "Q_VAN_XA"
   SymbolLibrary "Symbol library_101" at 857,824 size 9x40
      Appearance <- "Q_VAN_XA"
   SymbolLibrary "Symbol library_102" at 845,823 size 31x47
      Appearance <- "M_CB_CHAI"
   SymbolLibrary "Symbol library_103" at 411,126 size 47x31
      Appearance <- "M_CB_LOW_PG"
   SymbolLibrary "Symbol library_104" at 255,123 size 47x31
      Appearance <- "M_CB_LOW_MAU"
   SymbolLibrary "Symbol library_105" at 112,122 size 47x31
      Appearance <- "M_CB_LOW_HUONG"
   SymbolLibrary "Symbol library_106" at 520,168 size 47x31
      Appearance <- "M_CB_LOW_DUONG"
   SymbolLibrary "Symbol library_107" at 748,155 size 47x31
      Appearance <- "M_CB_LOW_NUOC"
   SymbolLibrary "Symbol library_108" at 972,141 size 47x31
      Appearance <- "M_CB_LOW_CO2"
   SymbolLibrary "Symbol library_109" at 564,933 size 59x70
      Appearance <- "Q_BT"
   SymbolLibrary "Symbol library_110" at 607,882 size 20x32
      Appearance <- "Q_VAN_XA"
      HorizontalMovement <- "TG_VT_SP"
   TextField "Text field_35" at 1333,93 size 170x24; Text 'BẢNG ĐIỀU KHIỂN'
   Switch "Switch_1" at 1282,129 size 100x54; TextOn 'AUTO'; CaptionText 'MODE'; TextOff 'MAN'
      on SwitchOff: ResetBit("M_mode")
      on SwitchOn: SetBit("M_mode")
      ProcessValue <- "M_mode"
   Button "Button_1" at 1282,191 size 96x32; TextOff 'Bắt Đầu'
      on Release: ResetBit("M_start")
      on Press: SetBit("M_start")
   Button "Button_2" at 1282,234 size 96x32; TextOff 'Dừng'
      on Release: ResetBit("M_Stop")
      on Press: SetBit("M_Stop")
   Circle "Circle_1" at 1413,143 size 48x48
      Appearance <- "Q_den_Auto"
   Circle "Circle_2" at 1500,143 size 48x48
      Appearance <- "Q_Den_Manual"
   Circle "Circle_3" at 1414,216 size 48x48
      Appearance <- "TG_DK_RUN"
   Circle "Circle_4" at 1497,218 size 48x48
      Appearance <- "Q_Den_loi"
   TextField "Text field_34" at 1417,156 size 38x18; Text 'AUTO'
   TextField "Text field_36" at 1507,157 size 33x18; Text 'MAN'
   TextField "Text field_37" at 1423,230 size 30x18; Text 'RUN'
   Switch "Switch_2" at 1283,266 size 100x54; TextOn 'ON'; CaptionText 'Mô Phỏng'; TextOff 'OFF'
      on SwitchOff: ResetBit("TG_Button_Simulation")
      on SwitchOn: SetBit("TG_Button_Simulation")
      ProcessValue <- "TG_Button_Simulation"
   TextField "Text field_38" at 1500,231 size 42x18; Text 'FAULT'
   TextField "Text field_39" at 1330,340 size 187x24; Text 'HIỂN THỊ THÔNG SỐ'
   TextField "Text field_40" at 1276,386 size 160x21; Text 'THỜI GIAN KHUẤY:'
   TextField "Text field_2" at 1278,414 size 138x21; Text 'NHIỆT ĐỘ TRỘN:'
   TextField "Text field_3" at 1281,444 size 117x21; Text 'NỒNG ĐỘ C02:'
   TextField "Text field_45" at 1291,505 size 240x24; Text 'HIỂN THỊ THÔNG SỐ MÁC'
   TextField "Text field_46" at 1259,546 size 211x21; Text 'TRỌNG LƯỢNG HƯƠNG VỊ:'
   TextField "Text field_4" at 1259,585 size 197x21; Text 'TRỌNG LƯỢNG PHỤ GIA:'
   TextField "Text field_5" at 1259,624 size 170x21; Text 'TRỌNG LƯỢNG MÀU:'
   TextField "Text field_6" at 1259,663 size 227x21; Text 'TRỌNG LƯỢNG NƯỚC TRỘN:'
   TextField "Text field_7" at 1259,702 size 213x21; Text 'TRỌNG LƯỢNG NƯỚC KHÍ:'
   TextField "Text field_8" at 1259,742 size 164x21; Text 'TRỌNG LƯỢNG CO2:'
   TextField "Text field_9" at 1309,826 size 230x24; Text 'THÔNG SỐ THÀNH PHẨM'
   TextField "Text field_10" at 1279,880 size 108x21; Text 'SẢN LƯỢNG :'
   TextField "Text field_11" at 1279,921 size 78x21; Text 'SỐ CHAI:'
   TextField "Text field_43" at 1553,389 size 23x21; Text '[S]'
   IOField "I/O field_14" at 1464,384 size 60x26; FormatPattern 9999999999
      ProcessValue <- "TL_thoiGian_khuay"
   IOField "I/O field_8" at 1464,415 size 60x26; FormatPattern 999.99
      ProcessValue <- "TL_nhietdo"
   IOField "I/O field_9" at 1464,446 size 60x26; FormatPattern 999.99
      ProcessValue <- "TL_CO2"
   IOField "I/O field_10" at 1487,551 size 60x26; FormatPattern 999.99
      ProcessValue <- "TL_Huong"
   IOField "I/O field_11" at 1487,588 size 60x26; FormatPattern 999.99
      ProcessValue <- "TL_PG"
   IOField "I/O field_12" at 1487,625 size 60x26; FormatPattern 999.99
      ProcessValue <- "TL_mau"
   IOField "I/O field_13" at 1487,663 size 60x26; FormatPattern 999.99
      ProcessValue <- "TL_nuoc_tron"
   IOField "I/O field_15" at 1487,700 size 60x26; FormatPattern 999.99
      ProcessValue <- "TL_Nuoc_KHi"
   IOField "I/O field_16" at 1487,738 size 60x26; FormatPattern 999.99
      ProcessValue <- "TL_CO2"
   IOField "I/O field_17" at 1424,879 size 60x26; FormatPattern 999.99
      ProcessValue <- "TL_San_Pham"
   IOField "I/O field_18" at 1424,915 size 60x26; FormatPattern 9999
      ProcessValue <- "Act_San_luong"
   TextField "Text field_28" at 1547,416 size 37x22; Text '[°C]'
   TextField "Text field_30" at 1546,445 size 40x27; Text '[g/l]'
   TextField "Text field_51" at 1549,553 size 38x21; Text '[KG]'
   TextField "Text field_12" at 1549,589 size 38x21; Text '[KG]'
   TextField "Text field_13" at 1549,626 size 38x21; Text '[KG]'
   TextField "Text field_14" at 1549,663 size 38x21; Text '[KG]'
   TextField "Text field_15" at 1549,701 size 38x21; Text '[KG]'
   TextField "Text field_16" at 1549,737 size 38x21; Text '[KG]'
   TextField "Text field_17" at 1527,876 size 38x21; Text '[KG]'
   Button "Button_6" at 101,213 size 58x28; TextOff 'V_H_1'
      on Release: ResetBit("M_SW_V1_Huong")
      on Press: SetBit("M_SW_V1_Huong")
   Button "Button_3" at 100,415 size 58x28; TextOff 'V_H_2'
      on Release: ResetBit("M_SW_V2_Huong")
      on Press: SetBit("M_SW_V2_Huong")
   Button "Button_4" at 252,212 size 58x28; TextOff 'V_M_1'
      on Release: ResetBit("M_SW_V1_mau")
      on Press: SetBit("M_SW_V1_mau")
   Button "Button_5" at 249,415 size 58x28; TextOff 'V_M_2'
      on Release: ResetBit("M_SW_V2_mau")
      on Press: SetBit("M_SW_V2_mau")
   Button "Button_7" at 390,415 size 58x28; TextOff 'V_PG_2'
      on Release: ResetBit("M_SW_V2_PG")
      on Press: SetBit("M_SW_V2_PG")
   Button "Button_8" at 524,415 size 58x28; TextOff 'V_D_2'
      on Release: ResetBit("M_SW_V2_Duong")
      on Press: SetBit("M_SW_V2_Duong")
   Button "Button_9" at 410,213 size 58x28; TextOff 'V_PG_1'
      on Release: ResetBit("M_SW_V1_PG")
      on Press: SetBit("M_SW_V1_PG")
   Button "Button_10" at 599,111 size 58x28; TextOff 'V_D_1'
      on Release: ResetBit("M_SW_V1_Duong")
      on Press: SetBit("M_SW_V1_Duong")
   Button "Button_11" at 603,274 size 58x28; TextOff 'V_NT_1'
      on Release: ResetBit("M_SW_V1_Nuoc_Tron")
      on Press: SetBit("M_SW_V1_Nuoc_Tron")
   Button "Button_12" at 809,190 size 58x28; TextOff 'V_NXK_1'
      on Release: ResetBit("M_SW_V1_Nuoc_Xuc_Khi")
      on Press: SetBit("M_SW_V1_Nuoc_Xuc_Khi")
   Button "Button_13" at 961,230 size 58x28; TextOff 'V_CO2_1'
      on Release: ResetBit("M_SW_V1_CO2")
      on Press: SetBit("M_SW_V1_CO2")
   Button "Button_14" at 957,428 size 58x28; TextOff 'V_CO2_2'
      on Release: ResetBit("M_SW_V2_CO2")
      on Press: SetBit("M_SW_V2_CO2")
   Button "Button_15" at 804,408 size 58x28; TextOff 'V_NXK_2'
      on Release: ResetBit("M_SW_V2_Nuoc_Xuc_Khi")
      on Press: SetBit("M_SW_V2_Nuoc_Xuc_Khi")
   Button "Button_16" at 682,400 size 58x28; TextOff 'V_NT_2'
      on Release: ResetBit("M_SW_V2_Nuoc_Tron")
      on Press: SetBit("M_SW_V2_Nuoc_Tron")
   Button "Button_17" at 373,557 size 58x28; TextOff 'TRON'
      on Release: ResetBit("M_SW_BOM_TRON")
      on Press: SetBit("M_SW_BOM_TRON")
   Button "Button_18" at 363,710 size 58x28; TextOff 'Bom_1'
      on Release: ResetBit("M_SW_BOM_1")
      on Press: SetBit("M_SW_BOM_1")
   Button "Button_19" at 773,702 size 58x28; TextOff 'Bom_2'
      on Release: ResetBit("M_SW_BOM_2")
      on Press: SetBit("M_SW_BOM_2")
   Button "Button_20" at 472,586 size 58x28; TextOff 'LANH'
      on Release: ResetBit("M_SW_LAM_LANH")
      on Press: SetBit("M_SW_LAM_LANH")
   Button "Button_21" at 915,756 size 58x28; TextOff 'V_X'
      on Release: ResetBit("M_SW_VAN_XA")
      on Press: SetBit("M_SW_VAN_XA")
   Button "Button_22" at 377,799 size 58x28; TextOff 'DOT'
      on Release: ResetBit("M_SW_LO_DOT")
      on Press: SetBit("M_SW_LO_DOT")
   TextField "Text field_18" at 43,70 size 87x42; Text 'HƯƠNG VỊ'
   TextField "Text field_19" at 204,70 size 47x23; Text 'MÀU'
   TextField "Text field_20" at 341,69 size 70x23; Text 'PHỤ GIA'
   TextField "Text field_21" at 454,74 size 66x23; Text 'ĐƯỜNG'
   TextField "Text field_22" at 700,53 size 53x23; Text 'NƯỚC'
   TextField "Text field_23" at 908,44 size 36x23; Text 'CO2'
   TextField "Text field_24" at 119,153 size 35x23; Text 'CB1'
   TextField "Text field_25" at 267,158 size 35x23; Text 'CB2'
   TextField "Text field_26" at 415,159 size 35x23; Text 'CB3'
   TextField "Text field_27" at 488,158 size 35x23; Text 'CB4'
   TextField "Text field_29" at 797,142 size 35x23; Text 'CB5'
   TextField "Text field_31" at 992,112 size 35x23; Text 'CB6'
   SymbolLibrary "Symbol library_111" at 558,541 size 31x47
      Appearance <- "M_CB_LOW_BON_2"
   TextField "Text field_32" at 520,529 size 35x23; Text 'CB8'
   TextField "Text field_33" at 814,824 size 35x23; Text 'CB8'
   TextField "Text field_41" at 102,184 size 94x23; Text 'Van Hương 1'
   TextField "Text field_42" at 247,184 size 79x23; Text 'Van Màu 1'
   TextField "Text field_44" at 406,189 size 68x23; Text 'Van PG 1'
   TextField "Text field_47" at 590,83 size 94x23; Text 'Van Đường 1'
   TextField "Text field_48" at 590,254 size 69x23; Text 'Van NT 1'
   TextField "Text field_49" at 796,224 size 82x23; Text 'Van NXK 1'
   TextField "Text field_50" at 956,207 size 78x23; Text 'Van CO2 1'
   TextField "Text field_52" at 97,390 size 94x23; Text 'Van Hương 2'
   TextField "Text field_53" at 248,389 size 79x23; Text 'Van Màu 2'
   TextField "Text field_54" at 389,389 size 68x23; Text 'Van PG 2'
   TextField "Text field_55" at 517,387 size 94x23; Text 'Van Đường 2'
   TextField "Text field_56" at 688,375 size 69x23; Text 'Van NT 2'
   TextField "Text field_57" at 808,380 size 82x23; Text 'Van NXK 2'
   TextField "Text field_58" at 951,392 size 78x23; Text 'Van CO2 1'
   TextField "Text field_59" at 376,591 size 72x23; Text 'Bơm Trộn'
   TextField "Text field_60" at 465,564 size 73x23; Text 'Làm Lạnh'
   TextField "Text field_61" at 367,737 size 49x23; Text 'Bơm 1'
   TextField "Text field_62" at 783,730 size 49x23; Text 'Bơm 2'
   TextField "Text field_63" at 381,772 size 52x23; Text 'Lò Đốt'
   TextField "Text field_64" at 912,730 size 58x23; Text 'Van_Xa'
   TextField "Text field_65" at 991,1 size 163x44; Text 'BẢNG DANH MỤC'
   Button "Button_23" at 1473,49 size 96x32; TextOff 'BIỂU ĐỒ>'; Authorization "Operate"
      on Press: ActivateScreen("Screen_2", 0)
   Button "Button_25" at 983,47 size 96x32; TextOff 'Đăng Xuất'
      on Activate: function_f23ef4c9(); ActivateScreen("DANG_NHAP", 0)
   Button "Button_26" at 1094,47 size 166x32; TextOff 'CÀI ĐẶT THÔNG SỐ'; Authorization "User administration"
      on Press: function_efd93a16("Cai_Dat_thong_So", 0, 0, -1, -1, 1)
   Button "Button_27" at 1282,48 size 166x32; TextOff 'CÀI ĐẶT MÁC'; Authorization "User administration"
      on Press: function_efd93a16("mac_tron", 0, 0, -1, -1, 1)
   TextField "Text field_66" at 109,262 size 83x23; Text 'Cân Hương'
   TextField "Text field_67" at 247,260 size 68x23; Text 'Cân Màu'
   TextField "Text field_68" at 398,251 size 89x23; Text 'Cân Phụ Gia'
   TextField "Text field_69" at 504,254 size 83x23; Text 'Cân Đường'
   TextField "Text field_70" at 685,250 size 92x23; Text 'Cân Nước_T'
   TextField "Text field_71" at 802,254 size 94x23; Text 'Cân Nước_K'
   TextField "Text field_72" at 961,260 size 67x23; Text 'Cân CO2'
   Button "Button_28" at 480,936 size 58x28; TextOff 'BT'
      on Release: ResetBit("M_SW_BANG_TAI")
      on Press: SetBit("M_SW_BANG_TAI")
   TextField "Text field_73" at 471,910 size 65x23; Text 'Bang Tai'
   TextField "Text field_74" at 1260,776 size 190x21; Text 'TRỌNG LƯỢNG ĐƯỜNG:'
   IOField "I/O field_19" at 1486,774 size 60x26; FormatPattern 999.99
      ProcessValue <- "TL_Duong"
   TextField "Text field_75" at 1550,774 size 38x21; Text '[KG]'
   TextField "Text field_76" at 1282,955 size 59x21; Text 'SỐ MẺ:'
   IOField "I/O field_20" at 1425,950 size 60x26; FormatPattern 99999
      ProcessValue <- "Act_me"
   IOField "I/O field_21" at 1405,3 size 166x40; FormatPattern ????????????????????????????????????????????????????????????????????????????????
      ProcessValue <- "Tag_Dang_nhap"
   SymbolLibrary "Symbol library_96" at 937,541 size 31x47
      Appearance <- "M_CB_LOW_BON_2"
   SymbolLibrary "Symbol library_112" at 337,540 size 31x47
      Appearance <- "M_CB_LOW_BON_2"
   TextField "Text field_77" at 944,512 size 35x23; Text 'CB9'
   TextField "Text field_78" at 366,526 size 35x23; Text 'CB7'

PopupScreen "mac_tron" 240x330
   Button "Button_2" at 16,11 size 201x32; TextOff 'Mác 150'
      on Press: SetTag("Set_Can_CO2", 30); SetTag("Set_can_Duong", 50); SetTag("Set_can_huong", 65); SetTag("Set_can_mau", 75); SetTag("Set_Can_nuoc_Tron", 50); SetTag("Set_Can_nuoc_xuc_khi", 40); SetTag("Set_can_PG", 80)
   Button "Button_1" at 16,58 size 199x32; TextOff 'Mác 200'
      on Press: SetTag("Set_Can_CO2", 40); SetTag("Set_can_Duong", 67); SetTag("Set_can_huong", 87); SetTag("Set_can_mau", 100); SetTag("Set_Can_nuoc_Tron", 67); SetTag("Set_Can_nuoc_xuc_khi", 53); SetTag("Set_can_PG", 107)
   Button "Button_3" at 16,119 size 198x32; TextOff 'Mác 250'
      on Press: SetTag("Set_Can_CO2", 50); SetTag("Set_can_Duong", 83); SetTag("Set_can_huong", 108); SetTag("Set_can_mau", 125); SetTag("Set_Can_nuoc_Tron", 83); SetTag("Set_Can_nuoc_xuc_khi", 67); SetTag("Set_can_PG", 133)
   Button "Button_4" at 16,172 size 196x32; TextOff 'Mác 300'
      on Press: SetTag("Set_Can_CO2", 60); SetTag("Set_can_Duong", 100); SetTag("Set_can_huong", 130); SetTag("Set_can_mau", 150); SetTag("Set_Can_nuoc_Tron", 100); SetTag("Set_Can_nuoc_xuc_khi", 80); SetTag("Set_can_PG", 160)
   Button "Button_5" at 16,222 size 196x32; TextOff 'Mác 350'
      on Press: SetTag("Set_Can_CO2", 70); SetTag("Set_can_Duong", 117); SetTag("Set_can_huong", 152); SetTag("Set_can_mau", 175); SetTag("Set_Can_nuoc_Tron", 117); SetTag("Set_Can_nuoc_xuc_khi", 93); SetTag("Set_can_PG", 187)
   Button "Button_6" at 16,276 size 196x32; TextOff 'Mác 400'
      on Press: SetTag("Set_Can_CO2", 80); SetTag("Set_can_Duong", 133); SetTag("Set_can_huong", 173); SetTag("Set_can_mau", 200); SetTag("Set_Can_nuoc_Tron", 133); SetTag("Set_Can_nuoc_xuc_khi", 107); SetTag("Set_can_PG", 213)

screen "Screen_2" 1600x1200
   TrendView "Trend view_1" at 43,69 size 1353x929
   Button "Button_1" at 1179,19 size 157x32; TextOff '<QUAY VỀ TRANG'
      on Press: ActivateScreen("Screen_1", 0)

PopupScreen "Cai_Dat_thong_So" 500x330
   TextField "Text field_39" at 131,14 size 180x24; Text 'CÀI ĐẶT THÔNG SỐ'
   TextField "Text field_40" at 11,54 size 192x21; Text 'SET THỜI GIAN KHUẤY:'
   TextField "Text field_1" at 11,79 size 71x21; Text 'SET MẺ:'
   TextField "Text field_2" at 11,110 size 122x21; Text 'SET NHIỆT ĐỘ:'
   TextField "Text field_3" at 11,137 size 210x21; Text 'SET KHỒI LƯỢNG HƯƠNG:'
   TextField "Text field_4" at 11,166 size 189x21; Text 'SET KHỒI LƯỢNG MÀU:'
   TextField "Text field_5" at 11,192 size 216x21; Text 'SET KHỒI LƯỢNG PHỤ GIA:'
   TextField "Text field_6" at 11,215 size 209x21; Text 'SET KHỒI LƯỢNG ĐƯỜNG:'
   TextField "Text field_7" at 11,243 size 246x21; Text 'SET KHỒI LƯỢNG NƯỚC TRỘN:'
   TextField "Text field_8" at 11,274 size 232x21; Text 'SET KHỒI LƯỢNG NƯỚC KHÍ:'
   TextField "Text field_9" at 11,303 size 233x21; Text 'SET KHỒI LƯỢNG NƯỚC CO2:'
   IOField "I/O field_14" at 332,49 size 60x26; FormatPattern 99999
      ProcessValue <- "Set_thoi_gian_khuay"
   IOField "I/O field_1" at 332,77 size 60x26; FormatPattern 99999
      ProcessValue <- "Set_me_tron"
   IOField "I/O field_2" at 332,105 size 60x26; FormatPattern 99999
      ProcessValue <- "Set_nhiet_do"
   IOField "I/O field_3" at 332,134 size 60x26; FormatPattern 99999
      ProcessValue <- "Set_can_huong"
   IOField "I/O field_4" at 332,163 size 60x26; FormatPattern 99999
      ProcessValue <- "Set_can_mau"
   IOField "I/O field_5" at 332,190 size 60x26; FormatPattern 99999
      ProcessValue <- "Set_can_PG"
   IOField "I/O field_6" at 332,217 size 60x26; FormatPattern 99999
      ProcessValue <- "Set_can_Duong"
   IOField "I/O field_7" at 332,244 size 60x26; FormatPattern 99999
      ProcessValue <- "Set_Can_nuoc_Tron"
   IOField "I/O field_8" at 332,273 size 60x26; FormatPattern 99999
      ProcessValue <- "Set_Can_nuoc_xuc_khi"
   IOField "I/O field_9" at 332,302 size 60x26; FormatPattern 99999
      ProcessValue <- "Set_Can_CO2"
   TextField "Text field_43" at 435,51 size 23x21; Text '[S]'
   TextField "Text field_28" at 435,107 size 37x22; Text '[°C]'
   TextField "Text field_30" at 435,302 size 40x27; Text '[g/l]'
   TextField "Text field_51" at 435,135 size 38x21; Text '[KG]'
   TextField "Text field_10" at 435,165 size 38x21; Text '[KG]'
   TextField "Text field_11" at 435,191 size 38x21; Text '[KG]'
   TextField "Text field_13" at 435,222 size 38x21; Text '[KG]'
   TextField "Text field_14" at 435,249 size 38x21; Text '[KG]'
   TextField "Text field_15" at 435,279 size 38x21; Text '[KG]'

screen "DANG_NHAP" 1600x1200
   GraphicView "Graphic view_1" at 0,0 size 1598x1198; Picture "Graphic_4"
   IOField "I/O field_1" at 575,408 size 324x54; FormatPattern ??????????????????????????????????????????????????
      ProcessValue <- "User_Input"
   IOField "I/O field_2" at 575,498 size 324x54; FormatPattern ??????????????????????????????????????????????????
      ProcessValue <- "Pass_Input"
   Button "Button_1" at 518,588 size 382x60; TextOff 'Đăng Nhập'
      on Click: function_a9b89908("Pass_Input", "User_Input")

VB script "LUU_CAI_DAT"
   On Error Resume Next
       Dim conn, sql
       Dim nguoiDung, setHuong, setMau, setPG, setDuong, setNT, setNK, setCO2, setMe, setTG, setNhiet
   
       ' 1. Đọc dữ liệu từ WinCC Tags (Đổi tên Tag trong ngoặc kép cho đúng với Project của bạn)
       nguoiDung = SmartTags("Tag_Dang_nhap")  ' Tag chứa tên người đăng nhập (Admin/User)
       setMe     = SmartTags("Set_me_tron")        ' Tên mác, VD: "Mác 150"
       setTG     = SmartTags("Set_thoi_gian_khuay")  ' Kiểu INT, không cần Replace
       
       ' Các tag kiểu FLOAT phải đổi dấu phẩy thành dấu chấm để SQL hiểu
       setHuong  = Replace(CStr(SmartTags("Set_can_huong")), ",", ".")
       setMau    = Replace(CStr(SmartTags("Set_can_mau")), ",", ".")
       setPG     = Replace(CStr(SmartTags("Set_can_PG")), ",", ".")
       setDuong  = Replace(CStr(SmartTags("Set_can_Duong")), ",", ".")
       setNT     = Replace(CStr(SmartTags("Set_Can_nuoc_Tron")), ",", ".")
       setNK     = Replace(CStr(SmartTags("Set_Can_nuoc_xuc_khi")), ",", ".")
       setCO2    = Replace(CStr(SmartTags("Set_Can_CO2")), ",", ".")
       setNhiet  = Replace(CStr(SmartTags("Set_nhiet_do")), ",", ".")
   
       ' 2. Mở kết nối ODBC
       Set conn = CreateObject("ADODB.Connection")
       conn.ConnectionString = "DSN=SYSTEM_WATER;"
       conn.Open
   
       ' 3. Thực thi câu lệnh SQL INSERT
       If conn.State = 1 Then
           sql = "INSERT INTO Bang_Cai_Dat (Nguoi_Truy_Cap, Set_Huong, Set_Mau, Set_Phu_Gia, Set_Duong, Set_Nuoc_Tron, Set_Nuoc_Khi, Set_CO2, Set_Me, Set_Thoi_Gian_Khuay, Set_Nhiet_Do) " & _
                 "VALUES ('" & nguoiDung & "', " & setHuong & ", " & setMau & ", " & setPG & ", " & setDuong & ", " & setNT & ", " & setNK & ", " & setCO2 & ", '" & setMe & "', " & setTG & ", " & setNhiet & ")"
           
           conn.Execute(sql)
           conn.Close
       End If
   
       Set conn = Nothing

VB script "LUU_GIA_TRI"
   On Error Resume Next
       Dim conn, sql
       Dim nguoiDung, huong, mau, duong, nuocTron, nuocKhi, co2, soMe, tgKhuay, nhietDo, soChai, tongTP
   
       ' 1. Đọc dữ liệu biến chuỗi
       nguoiDung = SmartTags("Tag_Dang_nhap")
       soMe      = SmartTags("Act_me")
       
       ' 2. Đọc dữ liệu số nguyên (INT)
       tgKhuay   = SmartTags("TL_thoiGian_khuay")
       soChai    = SmartTags("Act_San_luong") ' Chú ý: Hôm trước bạn gửi ảnh là Act_So_chai, hãy kiểm tra lại tên Tag này nhé!
   
       ' 3. Đọc và thay dấu phẩy thành dấu chấm cho biến FLOAT
       huong     = Replace(CStr(SmartTags("TL_Huong")), ",", ".")
       mau       = Replace(CStr(SmartTags("TL_mau")), ",", ".")
       duong     = Replace(CStr(SmartTags("TL_Duong")), ",", ".")
       nuocTron  = Replace(CStr(SmartTags("TL_nuoc_tron")), ",", ".")
       nuocKhi   = Replace(CStr(SmartTags("TL_Nuoc_KHi")), ",", ".")
       co2       = Replace(CStr(SmartTags("TL_CO2")), ",", ".")
       nhietDo   = Replace(CStr(SmartTags("TL_nhietdo")), ",", ".")
       tongTP    = Replace(CStr(SmartTags("TL_San_Pham")), ",", ".")
   
       Set conn = CreateObject("ADODB.Connection")
       conn.ConnectionString = "DSN=SYSTEM_WATER;"
       conn.Open
   
       ' 5. Thực thi câu lệnh SQL INSERT
       If conn.State = 1 Then
           sql = "INSERT INTO Bang_Thuc_Te (Nguoi_Truy_Cap, Khoi_Luong_Huong, Khoi_Luong_Mau, Khoi_Luong_Duong, Khoi_Luong_Nuoc_Tron, Khoi_Luong_Nuoc_Khi, Khoi_Luong_CO2, So_Me, Thoi_Gian_Khuay, Nhiet_Do, So_Chai, Tong_Thanh_Pham) " & _
                 "VALUES ('" & nguoiDung & "', " & huong & ", " & mau & ", " & duong & ", " & nuocTron & ", " & nuocKhi & ", " & co2 & ", '" & soMe & "', " & tgKhuay & ", " & nhietDo & ", " & soChai & ", " & tongTP & ")"
           
           conn.Execute(sql)
           conn.Close
       End If
   
       Set conn = Nothing

scheduled task "Get_user"
   on Action: function_f41c6f6c("Tag_Dang_nhap"); ActivateScreen("Screen_1", 0)

scheduled task "DATA_UPDATE_SETTING"
   Triggers <- "1 min"
   on Action: "LUU_CAI_DAT"('SYSTEM_WATER')

scheduled task "DATA_UPDATE_REAL"
   Triggers <- "1 min"
   on Action: "LUU_GIA_TRI"('SYSTEM_WATER')
*)